(* IEC 61131-3 sources: kns-pump-station/tests/POUs/Station/FB_StationCore_Test, 49 files *)

(* ---- AlarmIdCommandsResultAndClear.method.decl.st ---- *)
// 08 §14 вопрос 1: номера udiAckId, udiShelveId, udiUnshelveId — команда засчитывается, номер сбрасывается,
// результат — по ответу сводки
METHOD PRIVATE AlarmIdCommandsResultAndClear
VAR
    fbDut        : FB_StationCore;                    // ФБ под тестом
    fbTime       : PL.FB_FakeTime;                    // подменное время, старт 1 ч
    fbSink       : FB_FakeEventSink;                  // подменный журнал
    afbPump      : ARRAY[1..3] OF FB_FakeMotorVfd;    // подменные насосы: доступны, Auto, стоят
    stCmd        : ST_StationCmd;                     // GVL_Station.stStationCmd
    stCfgPersist : ST_StationCfg;                     // GVL_Persist.stStationCfg
    stCfgLkg     : ST_StationCfg;                     // GVL_Station.stCfgLkg
    stRetain     : ST_StationRetain;                  // GVL_Persist.stStationRetain
    fbPid        : PL.FB_PID;                         // GVL_Station.fbLIC101
    stPidCmd     : PL.ST_PidCmd;                      // GVL_Station.stLIC101Cmd
    stPidCfg     : PL.ST_PidCfg;                      // GVL_Persist.stLIC101Cfg
    stPidRetain  : PL.ST_DeviceRetain;                // GVL_Persist.stLIC101Retain
    fbAlarms     : FB_StationAlarms;                  // GVL_Station.fbAlarms
END_VAR

(* ---- ApplyProjectCfgChecksProjectLevelLimits.method.decl.st ---- *)
// 04 §18.3, DESIGN 6.15: «Применить уставки проекта» при LT101 L, перенастроенной наладчиком (1,1 м, станция —
// останов 1,2 м). PRG_Devices восстанавливает L/H LT101 уставок проекта в том же цикле, но после станции: уставки
// по умолчанию (останов 1,00 м) проверяются по L/H проекта (0,8 / 3,5 м). В цикле команды нет ложной ошибки уставок
// (NE 107 «функциональная проверка»), действующей становится копия по умолчанию, событие 101017 — одно, со значением 0
METHOD PRIVATE ApplyProjectCfgChecksProjectLevelLimits
VAR
    fbDut        : FB_StationCore;                    // ФБ под тестом
    fbTime       : PL.FB_FakeTime;                    // подменное время, старт 1 ч
    fbSink       : FB_FakeEventSink;                  // подменный журнал
    afbPump      : ARRAY[1..3] OF FB_FakeMotorVfd;    // подменные насосы: доступны, Auto, стоят
    stCmd        : ST_StationCmd;                     // GVL_Station.stStationCmd
    stCfgPersist : ST_StationCfg;                     // GVL_Persist.stStationCfg
    stCfgLkg     : ST_StationCfg;                     // GVL_Station.stCfgLkg
    stRetain     : ST_StationRetain;                  // GVL_Persist.stStationRetain
    fbPid        : PL.FB_PID;                         // GVL_Station.fbLIC101
    stPidCmd     : PL.ST_PidCmd;                      // GVL_Station.stLIC101Cmd
    stPidCfg     : PL.ST_PidCfg;                      // GVL_Persist.stLIC101Cfg
    stPidRetain  : PL.ST_DeviceRetain;                // GVL_Persist.stLIC101Retain
    fbAlarms     : FB_StationAlarms;                  // GVL_Station.fbAlarms
END_VAR

(* ---- ApplyProjectCfgRestoresDefaults.method.decl.st ---- *)
// 04 §18.3: «Применить уставки проекта» возвращает уставки станции и LIC101 к значениям GVL_StationDefaults
METHOD PRIVATE ApplyProjectCfgRestoresDefaults
VAR
    fbDut        : FB_StationCore;                    // ФБ под тестом
    fbTime       : PL.FB_FakeTime;                    // подменное время, старт 1 ч
    fbSink       : FB_FakeEventSink;                  // подменный журнал
    afbPump      : ARRAY[1..3] OF FB_FakeMotorVfd;    // подменные насосы: доступны, Auto, стоят
    stCmd        : ST_StationCmd;                     // GVL_Station.stStationCmd
    stCfgPersist : ST_StationCfg;                     // GVL_Persist.stStationCfg
    stCfgLkg     : ST_StationCfg;                     // GVL_Station.stCfgLkg
    stRetain     : ST_StationRetain;                  // GVL_Persist.stStationRetain
    fbPid        : PL.FB_PID;                         // GVL_Station.fbLIC101
    stPidCmd     : PL.ST_PidCmd;                      // GVL_Station.stLIC101Cmd
    stPidCfg     : PL.ST_PidCfg;                      // GVL_Persist.stLIC101Cfg
    stPidRetain  : PL.ST_DeviceRetain;                // GVL_Persist.stLIC101Retain
    fbAlarms     : FB_StationAlarms;                  // GVL_Station.fbAlarms
END_VAR

(* ---- AtsReplacesFaultedLead.method.decl.st ---- *)
// 04 §9, PMI-12, PMI-13: отказ ведущего — замена в том же цикле, событие 101006, KNS1.ATS
METHOD PRIVATE AtsReplacesFaultedLead
VAR
    fbDut        : FB_StationCore;                    // ФБ под тестом
    fbTime       : PL.FB_FakeTime;                    // подменное время, старт 1 ч
    fbSink       : FB_FakeEventSink;                  // подменный журнал
    afbPump      : ARRAY[1..3] OF FB_FakeMotorVfd;    // подменные насосы: доступны, Auto, стоят
    stCmd        : ST_StationCmd;                     // GVL_Station.stStationCmd
    stCfgPersist : ST_StationCfg;                     // GVL_Persist.stStationCfg
    stCfgLkg     : ST_StationCfg;                     // GVL_Station.stCfgLkg
    stRetain     : ST_StationRetain;                  // GVL_Persist.stStationRetain
    fbPid        : PL.FB_PID;                         // GVL_Station.fbLIC101
    stPidCmd     : PL.ST_PidCmd;                      // GVL_Station.stLIC101Cmd
    stPidCfg     : PL.ST_PidCfg;                      // GVL_Persist.stLIC101Cfg
    stPidRetain  : PL.ST_DeviceRetain;                // GVL_Persist.stLIC101Retain
    fbAlarms     : FB_StationAlarms;                  // GVL_Station.fbAlarms
END_VAR

(* ---- CommandPulsesClearedAndCounted.method.decl.st ---- *)
// 04 §19.2, контракт 2.1: импульсы и номера команд сбрасываются в том же цикле, uiCmdSeq растёт на число команд,
// eCmdResult — последней; события 101001, 101022, 101023
METHOD PRIVATE CommandPulsesClearedAndCounted
VAR
    fbDut        : FB_StationCore;                    // ФБ под тестом
    fbTime       : PL.FB_FakeTime;                    // подменное время, старт 1 ч
    fbSink       : FB_FakeEventSink;                  // подменный журнал
    afbPump      : ARRAY[1..3] OF FB_FakeMotorVfd;    // подменные насосы: доступны, Auto, стоят
    stCmd        : ST_StationCmd;                     // GVL_Station.stStationCmd
    stCfgPersist : ST_StationCfg;                     // GVL_Persist.stStationCfg
    stCfgLkg     : ST_StationCfg;                     // GVL_Station.stCfgLkg
    stRetain     : ST_StationRetain;                  // GVL_Persist.stStationRetain
    fbPid        : PL.FB_PID;                         // GVL_Station.fbLIC101
    stPidCmd     : PL.ST_PidCmd;                      // GVL_Station.stLIC101Cmd
    stPidCfg     : PL.ST_PidCfg;                      // GVL_Persist.stLIC101Cfg
    stPidRetain  : PL.ST_DeviceRetain;                // GVL_Persist.stLIC101Retain
    fbAlarms     : FB_StationAlarms;                  // GVL_Station.fbAlarms
    uiSeq0       : UINT;                              // счётчик команд до
END_VAR

(* ---- Cycle.method.decl.st ---- *)
// Помощник: uiSteps шагов времени tStep с вызовом ядра станции и всеми данными GVL_Station и
// GVL_Persist. xPlant — подменные насосы в Auto следуют запросам и общему заданию частоты
// (видно со следующего шага): работают, если запрошены, доступны и без отказа
METHOD PRIVATE Cycle
VAR_IN_OUT
    fbDut        : FB_StationCore;                    // ФБ под тестом
    fbTime       : PL.FB_FakeTime;                    // подменное время
    stCmd        : ST_StationCmd;                     // команды
    stCfgPersist : ST_StationCfg;                     // записанные уставки
    stCfgLkg     : ST_StationCfg;                     // действующая копия
    stRetain     : ST_StationRetain;                  // режим, способ
    fbPid        : PL.FB_PID;                         // LIC101
    stPidCmd     : PL.ST_PidCmd;                      // команды LIC101
    stPidCfg     : PL.ST_PidCfg;                      // уставки LIC101
    stPidRetain  : PL.ST_DeviceRetain;                // режим LIC101
    fbAlarms     : FB_StationAlarms;                  // тревоги станции
    afbPump      : ARRAY[1..3] OF FB_FakeMotorVfd;    // подменные насосы
END_VAR
VAR_INPUT
    tStep   : TIME;                                   // шаг времени
    uiSteps : UINT;                                   // шагов
    xPlant  : BOOL;                                   // насосы следуют запросам
END_VAR
VAR
    uiStep : UINT;                                    // номер шага
    uiIdx  : UINT;                                    // насос
END_VAR

(* ---- Cycle.method.impl.st ---- *)
FOR uiStep := 1 TO uiSteps DO
    fbTime.Advance(tStep := tStep);
    // сохранённая копия LKG — та же переменная, что и действующая: перезапуск ПЛК эти тесты не моделируют
    fbDut(itfTime := fbTime, stCmd := stCmd, stCfgPersist := stCfgPersist, stCfgLkg := stCfgLkg,
          stCfgLkgRetain := stCfgLkg, stRetain := stRetain, fbLIC101 := fbPid, stLIC101Cmd := stPidCmd,
          stLIC101Cfg := stPidCfg, stLIC101Retain := stPidRetain, fbAlarms := fbAlarms);
    IF xPlant THEN
        FOR uiIdx := 1 TO 3 DO
            IF afbPump[uiIdx].eMode = PL.E_DeviceMode.Auto THEN
                afbPump[uiIdx].xRunning := fbDut.axRun[uiIdx] AND afbPump[uiIdx].xAvailable
                                           AND NOT afbPump[uiIdx].xFault;
                afbPump[uiIdx].xSpeedAuto := afbPump[uiIdx].xRunning;
                afbPump[uiIdx].rSpeedRef := SEL(afbPump[uiIdx].xRunning, 0.0, fbDut.rSpeedSp_pct);
                afbPump[uiIdx].rSpeedAct := afbPump[uiIdx].rSpeedRef;
            END_IF
        END_FOR
    END_IF
END_FOR

(* ---- DryRunReleaseNoNoresStepFlicker.method.decl.st ---- *)
// 04 §7.4, §10.1, §15, PMI-22: выбран ПИД, сухой ход по LL дольше выдержек KNS1.NORES и KNS1.STEP (10 с) —
// обе подавлены (насосы заблокированы защитой станции). Насос видит снятие блокировки в своём вызове — после
// станции: в цикле снятия сухого хода насосы ещё недоступны, ПИД не готов. Ни NORES (High: сирена, K1), ни STEP
// не мелькают: выдержка появления отсчитывается заново после снятия подавления; затем снова ПИД
METHOD PRIVATE DryRunReleaseNoNoresStepFlicker
VAR
    fbDut        : FB_StationCore;                    // ФБ под тестом
    fbTime       : PL.FB_FakeTime;                    // подменное время, старт 1 ч
    fbSink       : FB_FakeEventSink;                  // подменный журнал
    afbPump      : ARRAY[1..3] OF FB_FakeMotorVfd;    // подменные насосы: доступны, Auto, стоят
    stCmd        : ST_StationCmd;                     // GVL_Station.stStationCmd
    stCfgPersist : ST_StationCfg;                     // GVL_Persist.stStationCfg
    stCfgLkg     : ST_StationCfg;                     // GVL_Station.stCfgLkg
    stRetain     : ST_StationRetain;                  // GVL_Persist.stStationRetain
    fbPid        : PL.FB_PID;                         // GVL_Station.fbLIC101
    stPidCmd     : PL.ST_PidCmd;                      // GVL_Station.stLIC101Cmd
    stPidCfg     : PL.ST_PidCfg;                      // GVL_Persist.stLIC101Cfg
    stPidRetain  : PL.ST_DeviceRetain;                // GVL_Persist.stLIC101Retain
    fbAlarms     : FB_StationAlarms;                  // GVL_Station.fbAlarms
    itfNores     : PL.I_Alarm;                        // KNS1.NORES через интерфейс
    itfStep      : PL.I_Alarm;                        // KNS1.STEP через интерфейс
    uiIdx        : UINT;                              // насос
    uiStep       : UINT;                              // шаг
    xFlicker     : BOOL;                              // NORES или STEP были неквитированными хотя бы в одном цикле
END_VAR

(* ---- DryRunReleaseNoNoresStepFlicker.method.impl.st ---- *)
coUnit.TEST('StationCore_DryRunReleaseNoNoresStepFlicker_A7_A10_A15_PMI22');

stPidCfg := GVL_StationDefaults.stLIC101Cfg;
stRetain.eMode := E_StationMode.Auto;
stRetain.eMethod := E_ControlMethod.LevelPid;
stPidRetain.eRemoteMode := PL.E_DeviceMode.Auto;
fbDut.aitfPump[1] := afbPump[1];
fbDut.aitfPump[2] := afbPump[2];
fbDut.aitfPump[3] := afbPump[3];
fbDut.axCommOk[1] := TRUE;
fbDut.axCommOk[2] := TRUE;
fbDut.axCommOk[3] := TRUE;
fbDut.itfEvents := fbSink;
fbDut.rLevel_m := 1.2;
fbDut.xLevelValid := TRUE;
fbDut.eLevelNe107 := PL.E_Ne107Status.Good;
fbDut.rLvlL_m := 0.8;
fbDut.rLvlH_m := 3.5;
fbDut.xPowerOk := TRUE;
Cycle(fbDut := fbDut, fbTime := fbTime, stCmd := stCmd, stCfgPersist := stCfgPersist, stCfgLkg := stCfgLkg,
      stRetain := stRetain, fbPid := fbPid, stPidCmd := stPidCmd, stPidCfg := stPidCfg,
      stPidRetain := stPidRetain, fbAlarms := fbAlarms, afbPump := afbPump, tStep := T#100MS, uiSteps := 110,
      xPlant := TRUE);

AssertTrue(Condition := fbDut.stSts.eControlAct = E_ControlAct.LevelPid, Message := 'LevelPid before dry run');
// LL по уровнемеру: сухой ход 20 с; насос недоступен с цикла после блокировки (как устройство после станции)
fbDut.rLevel_m := 0.45;
fbDut.xLevelL := TRUE;
fbDut.xLevelLL := TRUE;
FOR uiStep := 1 TO 200 DO
    Cycle(fbDut := fbDut, fbTime := fbTime, stCmd := stCmd, stCfgPersist := stCfgPersist, stCfgLkg := stCfgLkg,
          stRetain := stRetain, fbPid := fbPid, stPidCmd := stPidCmd, stPidCfg := stPidCfg,
          stPidRetain := stPidRetain, fbAlarms := fbAlarms, afbPump := afbPump, tStep := T#100MS, uiSteps := 1,
          xPlant := TRUE);
    FOR uiIdx := 1 TO 3 DO
        afbPump[uiIdx].xAvailable := fbDut.awInterlock[uiIdx] = 0;
    END_FOR
END_FOR

AssertTrue(Condition := fbDut.stSts.eControlAct = E_ControlAct.DryRunStop, Message := 'DryRunStop');
itfNores := fbAlarms.GetAlarm(uiIndex := E_StationAlarm.NORES - 1);
itfStep := fbAlarms.GetAlarm(uiIndex := E_StationAlarm.STEP - 1);
AssertTrue(Condition := itfNores.State = PL.E_AlarmState.SuppressedByDesign, Message := 'dry run: NORES suppressed');
AssertTrue(Condition := itfStep.State = PL.E_AlarmState.SuppressedByDesign, Message := 'dry run: STEP suppressed');
// уровень выше L: сухой ход снят
fbDut.rLevel_m := 1.0;
fbDut.xLevelL := FALSE;
fbDut.xLevelLL := FALSE;
xFlicker := FALSE;
FOR uiStep := 1 TO 150 DO
    Cycle(fbDut := fbDut, fbTime := fbTime, stCmd := stCmd, stCfgPersist := stCfgPersist, stCfgLkg := stCfgLkg,
          stRetain := stRetain, fbPid := fbPid, stPidCmd := stPidCmd, stPidCfg := stPidCfg,
          stPidRetain := stPidRetain, fbAlarms := fbAlarms, afbPump := afbPump, tStep := T#100MS, uiSteps := 1,
          xPlant := TRUE);
    IF uiStep = 1 THEN
        AssertEquals_UINT(Expected := 0, Actual := fbDut.stSts.uiPumpsAvailable,
                          Message := 'release cycle: pumps still interlocked');
    END_IF
    xFlicker := xFlicker OR (fbDut.stSts.wAlmUnack AND 16#0088) <> 0;
    FOR uiIdx := 1 TO 3 DO
        afbPump[uiIdx].xAvailable := fbDut.awInterlock[uiIdx] = 0;
    END_FOR
END_FOR

AssertFalse(Condition := xFlicker, Message := 'no unacked KNS1.NORES or KNS1.STEP on dry run release');
AssertTrue(Condition := itfNores.State = PL.E_AlarmState.Normal, Message := 'NORES normal');
AssertTrue(Condition := itfStep.State = PL.E_AlarmState.Normal, Message := 'STEP normal');
AssertTrue(Condition := fbDut.stSts.eControlAct = E_ControlAct.LevelPid, Message := 'LevelPid after dry run');

coUnit.TEST_FINISHED();

(* ---- DryRunStopSuppressesNoReserve.method.decl.st ---- *)
// 04 §10.1, §11, §15, PMI-21: откачка по поплавкам до LS103 — сухой ход блокирует все насосы (Available = FALSE).
// Насосы стоят по защите станции, а не из-за отказов: KNS1.NORES подавлена (дубль KNS1.DRY, иначе High-тревога и
// обесточенное K1 в каждом цикле откачки по поплавкам)
METHOD PRIVATE DryRunStopSuppressesNoReserve
VAR
    fbDut        : FB_StationCore;                    // ФБ под тестом
    fbTime       : PL.FB_FakeTime;                    // подменное время, старт 1 ч
    fbSink       : FB_FakeEventSink;                  // подменный журнал
    afbPump      : ARRAY[1..3] OF FB_FakeMotorVfd;    // подменные насосы: доступны, Auto, стоят
    stCmd        : ST_StationCmd;                     // GVL_Station.stStationCmd
    stCfgPersist : ST_StationCfg;                     // GVL_Persist.stStationCfg
    stCfgLkg     : ST_StationCfg;                     // GVL_Station.stCfgLkg
    stRetain     : ST_StationRetain;                  // GVL_Persist.stStationRetain
    fbPid        : PL.FB_PID;                         // GVL_Station.fbLIC101
    stPidCmd     : PL.ST_PidCmd;                      // GVL_Station.stLIC101Cmd
    stPidCfg     : PL.ST_PidCfg;                      // GVL_Persist.stLIC101Cfg
    stPidRetain  : PL.ST_DeviceRetain;                // GVL_Persist.stLIC101Retain
    fbAlarms     : FB_StationAlarms;                  // GVL_Station.fbAlarms
    itfAlm       : PL.I_Alarm;                        // тревога через интерфейс
    uiIdx        : UINT;                              // насос
END_VAR

(* ---- DryRunStopSuppressesNoReserve.method.impl.st ---- *)
coUnit.TEST('StationCore_DryRunStopSuppressesNoReserve_A10_A11_A15_PMI21');

stPidCfg := GVL_StationDefaults.stLIC101Cfg;
stRetain.eMode := E_StationMode.Auto;
fbDut.aitfPump[1] := afbPump[1];
fbDut.aitfPump[2] := afbPump[2];
fbDut.aitfPump[3] := afbPump[3];
fbDut.axCommOk[1] := TRUE;
fbDut.axCommOk[2] := TRUE;
fbDut.axCommOk[3] := TRUE;
fbDut.itfEvents := fbSink;
fbDut.rLevel_m := 1.2;
fbDut.xLevelValid := TRUE;
fbDut.eLevelNe107 := PL.E_Ne107Status.Good;
fbDut.rLvlL_m := 0.8;
fbDut.rLvlH_m := 3.5;
fbDut.xPowerOk := TRUE;
Cycle(fbDut := fbDut, fbTime := fbTime, stCmd := stCmd, stCfgPersist := stCfgPersist, stCfgLkg := stCfgLkg,
      stRetain := stRetain, fbPid := fbPid, stPidCmd := stPidCmd, stPidCfg := stPidCfg,
      stPidRetain := stPidRetain, fbAlarms := fbAlarms, afbPump := afbPump, tStep := T#100MS, uiSteps := 110,
      xPlant := TRUE);

// отказ LT101, LS102: откачка всеми насосами
fbDut.xLevelValid := FALSE;
fbDut.xFloatHigh := TRUE;
Cycle(fbDut := fbDut, fbTime := fbTime, stCmd := stCmd, stCfgPersist := stCfgPersist, stCfgLkg := stCfgLkg,
      stRetain := stRetain, fbPid := fbPid, stPidCmd := stPidCmd, stPidCfg := stPidCfg,
      stPidRetain := stPidRetain, fbAlarms := fbAlarms, afbPump := afbPump, tStep := T#100MS, uiSteps := 110,
      xPlant := TRUE);

AssertTrue(Condition := afbPump[1].xRunning AND afbPump[2].xRunning AND afbPump[3].xRunning, Message := 'pumping');
// уровень у LS103: сухой ход, блокировка всех насосов — устройства недоступны и стоят
fbDut.xFloatHigh := FALSE;
fbDut.xFloatDry := TRUE;
Cycle(fbDut := fbDut, fbTime := fbTime, stCmd := stCmd, stCfgPersist := stCfgPersist, stCfgLkg := stCfgLkg,
      stRetain := stRetain, fbPid := fbPid, stPidCmd := stPidCmd, stPidCfg := stPidCfg,
      stPidRetain := stPidRetain, fbAlarms := fbAlarms, afbPump := afbPump, tStep := T#100MS, uiSteps := 1,
      xPlant := TRUE);

AssertTrue(Condition := (fbDut.awInterlock[1] AND GVL_Const.KNS_ILK_DRY_RUN) <> 0, Message := 'dry run interlock');
FOR uiIdx := 1 TO 3 DO
    afbPump[uiIdx].xAvailable := FALSE;
END_FOR
Cycle(fbDut := fbDut, fbTime := fbTime, stCmd := stCmd, stCfgPersist := stCfgPersist, stCfgLkg := stCfgLkg,
      stRetain := stRetain, fbPid := fbPid, stPidCmd := stPidCmd, stPidCfg := stPidCfg,
      stPidRetain := stPidRetain, fbAlarms := fbAlarms, afbPump := afbPump, tStep := T#100MS, uiSteps := 200,
      xPlant := TRUE);

AssertTrue(Condition := fbDut.stSts.eControlAct = E_ControlAct.DryRunStop, Message := 'DryRunStop');
AssertEquals_UINT(Expected := 0, Actual := fbDut.stSts.uiPumpsAvailable, Message := 'no pump available');
itfAlm := fbAlarms.GetAlarm(uiIndex := E_StationAlarm.NORES - 1);
AssertTrue(Condition := itfAlm.State = PL.E_AlarmState.SuppressedByDesign, Message := 'NORES suppressed by dry run');
AssertEquals_WORD(Expected := 0, Actual := fbDut.stSts.wAlmActive AND 16#0004, Message := 'no LACK');
AssertEquals_WORD(Expected := 0, Actual := fbDut.stSts.wAlmUnack AND 16#000C, Message := 'no LACK, NORES unacked');
AssertEquals_WORD(Expected := 0, Actual := fbDut.stSts.wState AND GVL_Const.STN_ST_NO_RESERVE,
                  Message := 'wState: no reserve bit clear');

coUnit.TEST_FINISHED();

(* ---- EmergencyRequiresAllAtFullSpeed.method.decl.st ---- *)
// 04 §10.2, PMI-20: аварийный уровень в «Автомате» — требуются все три насоса, задание 100 %, KNS1.EHL, K1 по
// сводке
METHOD PRIVATE EmergencyRequiresAllAtFullSpeed
VAR
    fbDut        : FB_StationCore;                    // ФБ под тестом
    fbTime       : PL.FB_FakeTime;                    // подменное время, старт 1 ч
    fbSink       : FB_FakeEventSink;                  // подменный журнал
    afbPump      : ARRAY[1..3] OF FB_FakeMotorVfd;    // подменные насосы: доступны, Auto, стоят
    stCmd        : ST_StationCmd;                     // GVL_Station.stStationCmd
    stCfgPersist : ST_StationCfg;                     // GVL_Persist.stStationCfg
    stCfgLkg     : ST_StationCfg;                     // GVL_Station.stCfgLkg
    stRetain     : ST_StationRetain;                  // GVL_Persist.stStationRetain
    fbPid        : PL.FB_PID;                         // GVL_Station.fbLIC101
    stPidCmd     : PL.ST_PidCmd;                      // GVL_Station.stLIC101Cmd
    stPidCfg     : PL.ST_PidCfg;                      // GVL_Persist.stLIC101Cfg
    stPidRetain  : PL.ST_DeviceRetain;                // GVL_Persist.stLIC101Retain
    fbAlarms     : FB_StationAlarms;                  // GVL_Station.fbAlarms
END_VAR

(* ---- ExportCommandAndEvents.method.decl.st ---- *)
// 04 §16, PMI-37: xExportLog — запрос снимка; во время выгрузки отклоняется; переход в Done — событие 101019 с
// числом строк, в Error — 101020
METHOD PRIVATE ExportCommandAndEvents
VAR
    fbDut        : FB_StationCore;                    // ФБ под тестом
    fbTime       : PL.FB_FakeTime;                    // подменное время, старт 1 ч
    fbSink       : FB_FakeEventSink;                  // подменный журнал
    afbPump      : ARRAY[1..3] OF FB_FakeMotorVfd;    // подменные насосы: доступны, Auto, стоят
    stCmd        : ST_StationCmd;                     // GVL_Station.stStationCmd
    stCfgPersist : ST_StationCfg;                     // GVL_Persist.stStationCfg
    stCfgLkg     : ST_StationCfg;                     // GVL_Station.stCfgLkg
    stRetain     : ST_StationRetain;                  // GVL_Persist.stStationRetain
    fbPid        : PL.FB_PID;                         // GVL_Station.fbLIC101
    stPidCmd     : PL.ST_PidCmd;                      // GVL_Station.stLIC101Cmd
    stPidCfg     : PL.ST_PidCfg;                      // GVL_Persist.stLIC101Cfg
    stPidRetain  : PL.ST_DeviceRetain;                // GVL_Persist.stLIC101Retain
    fbAlarms     : FB_StationAlarms;                  // GVL_Station.fbAlarms
END_VAR

(* ---- FloatModeStartsAllOnLs102.method.decl.st ---- *)
// 04 §11, PMI-21, PMI-25: LT101 недостоверен — Float; LS102 — все насосы, 100 %; KNS1.EHL и KNS1.DRY подавлены,
// KNS1.FLOAT активна
METHOD PRIVATE FloatModeStartsAllOnLs102
VAR
    fbDut        : FB_StationCore;                    // ФБ под тестом
    fbTime       : PL.FB_FakeTime;                    // подменное время, старт 1 ч
    fbSink       : FB_FakeEventSink;                  // подменный журнал
    afbPump      : ARRAY[1..3] OF FB_FakeMotorVfd;    // подменные насосы: доступны, Auto, стоят
    stCmd        : ST_StationCmd;                     // GVL_Station.stStationCmd
    stCfgPersist : ST_StationCfg;                     // GVL_Persist.stStationCfg
    stCfgLkg     : ST_StationCfg;                     // GVL_Station.stCfgLkg
    stRetain     : ST_StationRetain;                  // GVL_Persist.stStationRetain
    fbPid        : PL.FB_PID;                         // GVL_Station.fbLIC101
    stPidCmd     : PL.ST_PidCmd;                      // GVL_Station.stLIC101Cmd
    stPidCfg     : PL.ST_PidCfg;                      // GVL_Persist.stLIC101Cfg
    stPidRetain  : PL.ST_DeviceRetain;                // GVL_Persist.stLIC101Retain
    fbAlarms     : FB_StationAlarms;                  // GVL_Station.fbAlarms
    itfAlm       : PL.I_Alarm;                        // тревога через интерфейс
END_VAR

(* ---- FlowAlarmsSuppressedUntilSettled.method.decl.st ---- *)
// DESIGN 7, шаг 12: тревоги L/LL PT201 и L FT202 подавлены, пока ни один насос не работает дольше STN_FLOW_SETTLE
// = 20 с
METHOD PRIVATE FlowAlarmsSuppressedUntilSettled
VAR
    fbDut        : FB_StationCore;                    // ФБ под тестом
    fbTime       : PL.FB_FakeTime;                    // подменное время, старт 1 ч
    fbSink       : FB_FakeEventSink;                  // подменный журнал
    afbPump      : ARRAY[1..3] OF FB_FakeMotorVfd;    // подменные насосы: доступны, Auto, стоят
    stCmd        : ST_StationCmd;                     // GVL_Station.stStationCmd
    stCfgPersist : ST_StationCfg;                     // GVL_Persist.stStationCfg
    stCfgLkg     : ST_StationCfg;                     // GVL_Station.stCfgLkg
    stRetain     : ST_StationRetain;                  // GVL_Persist.stStationRetain
    fbPid        : PL.FB_PID;                         // GVL_Station.fbLIC101
    stPidCmd     : PL.ST_PidCmd;                      // GVL_Station.stLIC101Cmd
    stPidCfg     : PL.ST_PidCfg;                      // GVL_Persist.stLIC101Cfg
    stPidRetain  : PL.ST_DeviceRetain;                // GVL_Persist.stLIC101Retain
    fbAlarms     : FB_StationAlarms;                  // GVL_Station.fbAlarms
END_VAR

(* ---- LackSuppressesNoReserve.method.decl.st ---- *)
// 04 §15, PMI-17: недостаточно насосов — KNS1.LACK через 10 с, KNS1.NORES подавлена; NE 107 станции — Failure
METHOD PRIVATE LackSuppressesNoReserve
VAR
    fbDut        : FB_StationCore;                    // ФБ под тестом
    fbTime       : PL.FB_FakeTime;                    // подменное время, старт 1 ч
    fbSink       : FB_FakeEventSink;                  // подменный журнал
    afbPump      : ARRAY[1..3] OF FB_FakeMotorVfd;    // подменные насосы: доступны, Auto, стоят
    stCmd        : ST_StationCmd;                     // GVL_Station.stStationCmd
    stCfgPersist : ST_StationCfg;                     // GVL_Persist.stStationCfg
    stCfgLkg     : ST_StationCfg;                     // GVL_Station.stCfgLkg
    stRetain     : ST_StationRetain;                  // GVL_Persist.stStationRetain
    fbPid        : PL.FB_PID;                         // GVL_Station.fbLIC101
    stPidCmd     : PL.ST_PidCmd;                      // GVL_Station.stLIC101Cmd
    stPidCfg     : PL.ST_PidCfg;                      // GVL_Persist.stLIC101Cfg
    stPidRetain  : PL.ST_DeviceRetain;                // GVL_Persist.stLIC101Retain
    fbAlarms     : FB_StationAlarms;                  // GVL_Station.fbAlarms
    itfAlm       : PL.I_Alarm;                        // тревога через интерфейс
END_VAR

(* ---- LkgRejectsInvalidCfg.method.decl.st ---- *)
// 04 §18.3, PMI-08: корректная уставка принимается (событие 101017 с номером параметра 8), неверная не применяется
// — бит wCfgErr, работа по последней корректной копии
METHOD PRIVATE LkgRejectsInvalidCfg
VAR
    fbDut        : FB_StationCore;                    // ФБ под тестом
    fbTime       : PL.FB_FakeTime;                    // подменное время, старт 1 ч
    fbSink       : FB_FakeEventSink;                  // подменный журнал
    afbPump      : ARRAY[1..3] OF FB_FakeMotorVfd;    // подменные насосы: доступны, Auto, стоят
    stCmd        : ST_StationCmd;                     // GVL_Station.stStationCmd
    stCfgPersist : ST_StationCfg;                     // GVL_Persist.stStationCfg
    stCfgLkg     : ST_StationCfg;                     // GVL_Station.stCfgLkg
    stRetain     : ST_StationRetain;                  // GVL_Persist.stStationRetain
    fbPid        : PL.FB_PID;                         // GVL_Station.fbLIC101
    stPidCmd     : PL.ST_PidCmd;                      // GVL_Station.stLIC101Cmd
    stPidCfg     : PL.ST_PidCfg;                      // GVL_Persist.stLIC101Cfg
    stPidRetain  : PL.ST_DeviceRetain;                // GVL_Persist.stLIC101Retain
    fbAlarms     : FB_StationAlarms;                  // GVL_Station.fbAlarms
END_VAR

(* ---- LkgRestoredAfterRestart.method.decl.st ---- *)
// 04 §18.3, PMI-08, PMI-35: последняя корректная копия уставок переживает перезапуск ПЛК. Корректная правка
// (задание 1,8 м) принята и сохранена в энергонезависимой копии LKG, неверная (2,5 м) осталась в записанных
// уставках; после перезапуска (новый экземпляр ядра, GVL_Station.stCfgLkg — умолчания) станция работает по
// сохранённой копии 1,8 м, а не по уставкам проекта; событие 101017 при старте не пишется
METHOD PRIVATE LkgRestoredAfterRestart
VAR
    fbTime         : PL.FB_FakeTime;                  // подменное время, старт 1 ч
    afbPump        : ARRAY[1..3] OF FB_FakeMotorVfd;  // подменные насосы: доступны, Auto, стоят
    // энергонезависимые данные (GVL_Persist): переживают перезапуск
    stCfgPersist   : ST_StationCfg;                   // GVL_Persist.stStationCfg
    stCfgLkgRetain : ST_StationCfg;                   // GVL_Persist.stStationCfgLkg
    stRetain       : ST_StationRetain;                // GVL_Persist.stStationRetain
    stPidCfg       : PL.ST_PidCfg;                    // GVL_Persist.stLIC101Cfg
    stPidRetain    : PL.ST_DeviceRetain;              // GVL_Persist.stLIC101Retain
END_VAR
VAR_INST
    // до перезапуска
    fbDutBefore    : FB_StationCore;                  // ядро до перезапуска
    fbSinkBefore   : FB_FakeEventSink;                // журнал до перезапуска
    stCmdBefore    : ST_StationCmd;                   // GVL_Station.stStationCmd
    stLkgBefore    : ST_StationCfg;                   // GVL_Station.stCfgLkg
    fbPidBefore    : PL.FB_PID;                       // GVL_Station.fbLIC101
    stPidCmdBefore : PL.ST_PidCmd;                    // GVL_Station.stLIC101Cmd
    fbAlmBefore    : FB_StationAlarms;                // GVL_Station.fbAlarms
    // после перезапуска: обычные переменные снова с умолчаниями
    fbDutAfter     : FB_StationCore;                  // ядро после перезапуска
    fbSinkAfter    : FB_FakeEventSink;                // журнал после перезапуска
    stCmdAfter     : ST_StationCmd;
    stLkgAfter     : ST_StationCfg;
    fbPidAfter     : PL.FB_PID;
    stPidCmdAfter  : PL.ST_PidCmd;
    fbAlmAfter     : FB_StationAlarms;
END_VAR

(* ---- ManualDryRunInterlocksAllPumps.method.decl.st ---- *)
// 04 §10.1, PMI-18: в «Ручном» запросов нет, но сухой ход по LL блокирует все насосы (KNS_ILK_DRY_RUN), тревога
// KNS1.DRY
METHOD PRIVATE ManualDryRunInterlocksAllPumps
VAR
    fbDut        : FB_StationCore;                    // ФБ под тестом
    fbTime       : PL.FB_FakeTime;                    // подменное время, старт 1 ч
    fbSink       : FB_FakeEventSink;                  // подменный журнал
    afbPump      : ARRAY[1..3] OF FB_FakeMotorVfd;    // подменные насосы: доступны, Auto, стоят
    stCmd        : ST_StationCmd;                     // GVL_Station.stStationCmd
    stCfgPersist : ST_StationCfg;                     // GVL_Persist.stStationCfg
    stCfgLkg     : ST_StationCfg;                     // GVL_Station.stCfgLkg
    stRetain     : ST_StationRetain;                  // GVL_Persist.stStationRetain
    fbPid        : PL.FB_PID;                         // GVL_Station.fbLIC101
    stPidCmd     : PL.ST_PidCmd;                      // GVL_Station.stLIC101Cmd
    stPidCfg     : PL.ST_PidCfg;                      // GVL_Persist.stLIC101Cfg
    stPidRetain  : PL.ST_DeviceRetain;                // GVL_Persist.stLIC101Retain
    fbAlarms     : FB_StationAlarms;                  // GVL_Station.fbAlarms
END_VAR

(* ---- ManualFloatModeKeepsEhlDry.method.decl.st ---- *)
// 04 §3.1, §10.2, §11, §15: станция в «Ручном», LT101 отказал. Управления по поплавкам в «Ручном» нет (насосы
// автоматика не пускает), поэтому KNS1.EHL (Critical) по LS102 и KNS1.DRY по LS103 не подавляются: подавление
// «режим по поплавкам» действует только в «Автомате», где срабатывания поплавков — штатные точки управления
METHOD PRIVATE ManualFloatModeKeepsEhlDry
VAR
    fbDut        : FB_StationCore;                    // ФБ под тестом
    fbTime       : PL.FB_FakeTime;                    // подменное время, старт 1 ч
    fbSink       : FB_FakeEventSink;                  // подменный журнал
    afbPump      : ARRAY[1..3] OF FB_FakeMotorVfd;    // подменные насосы: доступны, Auto, стоят
    stCmd        : ST_StationCmd;                     // GVL_Station.stStationCmd
    stCfgPersist : ST_StationCfg;                     // GVL_Persist.stStationCfg
    stCfgLkg     : ST_StationCfg;                     // GVL_Station.stCfgLkg
    stRetain     : ST_StationRetain;                  // GVL_Persist.stStationRetain
    fbPid        : PL.FB_PID;                         // GVL_Station.fbLIC101
    stPidCmd     : PL.ST_PidCmd;                      // GVL_Station.stLIC101Cmd
    stPidCfg     : PL.ST_PidCfg;                      // GVL_Persist.stLIC101Cfg
    stPidRetain  : PL.ST_DeviceRetain;                // GVL_Persist.stLIC101Retain
    fbAlarms     : FB_StationAlarms;                  // GVL_Station.fbAlarms
    itfEhl       : PL.I_Alarm;                        // KNS1.EHL через интерфейс
    itfDry       : PL.I_Alarm;                        // KNS1.DRY через интерфейс
END_VAR

(* ---- ManualToAutoAdoptsRunningPump.method.decl.st ---- *)
// 04 §3.2, PMI-30: «Ручной» → «Автомат» при работающем насосе — в том же цикле запрос ему (без останова), насосам
// — RequestMode(Auto), задание частоты следило за насосом
METHOD PRIVATE ManualToAutoAdoptsRunningPump
VAR
    fbDut        : FB_StationCore;                    // ФБ под тестом
    fbTime       : PL.FB_FakeTime;                    // подменное время, старт 1 ч
    fbSink       : FB_FakeEventSink;                  // подменный журнал
    afbPump      : ARRAY[1..3] OF FB_FakeMotorVfd;    // подменные насосы: доступны, Auto, стоят
    stCmd        : ST_StationCmd;                     // GVL_Station.stStationCmd
    stCfgPersist : ST_StationCfg;                     // GVL_Persist.stStationCfg
    stCfgLkg     : ST_StationCfg;                     // GVL_Station.stCfgLkg
    stRetain     : ST_StationRetain;                  // GVL_Persist.stStationRetain
    fbPid        : PL.FB_PID;                         // GVL_Station.fbLIC101
    stPidCmd     : PL.ST_PidCmd;                      // GVL_Station.stLIC101Cmd
    stPidCfg     : PL.ST_PidCfg;                      // GVL_Persist.stLIC101Cfg
    stPidRetain  : PL.ST_DeviceRetain;                // GVL_Persist.stLIC101Retain
    fbAlarms     : FB_StationAlarms;                  // GVL_Station.fbAlarms
END_VAR

(* ---- ManualToAutoStoppedPumpsNoNoresFlicker.method.decl.st ---- *)
// 04 §3.2, §15, PMI-30: «Ручной» дольше выдержки KNS1.NORES (10 с) при остановленных насосах, затем «Автомат».
// Насос выполняет запрос режима в своём вызове — после станции: в цикле входа в «Автомат» насосы ещё в Manual
// (доступных нет), подавление «Ручной» уже снято, а требуемое число 0 (KNS1.LACK нет). Тревога не мелькает
// (High: сирена, K1): выдержка появления отсчитывается заново после снятия подавления
METHOD PRIVATE ManualToAutoStoppedPumpsNoNoresFlicker
VAR
    fbDut        : FB_StationCore;                    // ФБ под тестом
    fbTime       : PL.FB_FakeTime;                    // подменное время, старт 1 ч
    fbSink       : FB_FakeEventSink;                  // подменный журнал
    afbPump      : ARRAY[1..3] OF FB_FakeMotorVfd;    // подменные насосы: доступны, Auto, стоят
    stCmd        : ST_StationCmd;                     // GVL_Station.stStationCmd
    stCfgPersist : ST_StationCfg;                     // GVL_Persist.stStationCfg
    stCfgLkg     : ST_StationCfg;                     // GVL_Station.stCfgLkg
    stRetain     : ST_StationRetain;                  // GVL_Persist.stStationRetain
    fbPid        : PL.FB_PID;                         // GVL_Station.fbLIC101
    stPidCmd     : PL.ST_PidCmd;                      // GVL_Station.stLIC101Cmd
    stPidCfg     : PL.ST_PidCfg;                      // GVL_Persist.stLIC101Cfg
    stPidRetain  : PL.ST_DeviceRetain;                // GVL_Persist.stLIC101Retain
    fbAlarms     : FB_StationAlarms;                  // GVL_Station.fbAlarms
    itfAlm       : PL.I_Alarm;                        // KNS1.NORES через интерфейс
    uiIdx        : UINT;                              // насос
    uiStep       : UINT;                              // шаг
    xFlicker     : BOOL;                              // NORES была неквитированной хотя бы в одном цикле
END_VAR

(* ---- ManualToAutoStoppedPumpsNoNoresFlicker.method.impl.st ---- *)
coUnit.TEST('StationCore_ManualToAutoStoppedPumpsNoNoresFlicker_A3_A15_PMI30');

stPidCfg := GVL_StationDefaults.stLIC101Cfg;
stRetain.eMode := E_StationMode.Auto;
fbDut.aitfPump[1] := afbPump[1];
fbDut.aitfPump[2] := afbPump[2];
fbDut.aitfPump[3] := afbPump[3];
fbDut.axCommOk[1] := TRUE;
fbDut.axCommOk[2] := TRUE;
fbDut.axCommOk[3] := TRUE;
fbDut.itfEvents := fbSink;
fbDut.rLevel_m := 1.2;
fbDut.xLevelValid := TRUE;
fbDut.eLevelNe107 := PL.E_Ne107Status.Good;
fbDut.rLvlL_m := 0.8;
fbDut.rLvlH_m := 3.5;
fbDut.xPowerOk := TRUE;
Cycle(fbDut := fbDut, fbTime := fbTime, stCmd := stCmd, stCfgPersist := stCfgPersist, stCfgLkg := stCfgLkg,
      stRetain := stRetain, fbPid := fbPid, stPidCmd := stPidCmd, stPidCfg := stPidCfg,
      stPidRetain := stPidRetain, fbAlarms := fbAlarms, afbPump := afbPump, tStep := T#100MS, uiSteps := 110,
      xPlant := TRUE);

// «Ручной»: насосы выполняют запрос в своём вызове (циклом позже станции)
stCmd.xSetManual := TRUE;
Cycle(fbDut := fbDut, fbTime := fbTime, stCmd := stCmd, stCfgPersist := stCfgPersist, stCfgLkg := stCfgLkg,
      stRetain := stRetain, fbPid := fbPid, stPidCmd := stPidCmd, stPidCfg := stPidCfg,
      stPidRetain := stPidRetain, fbAlarms := fbAlarms, afbPump := afbPump, tStep := T#100MS, uiSteps := 1,
      xPlant := TRUE);

FOR uiIdx := 1 TO 3 DO
    afbPump[uiIdx].eMode := afbPump[uiIdx].eLastModeRequest;
END_FOR
AssertTrue(Condition := afbPump[1].eMode = PL.E_DeviceMode.Manual, Message := 'pumps in Manual');
Cycle(fbDut := fbDut, fbTime := fbTime, stCmd := stCmd, stCfgPersist := stCfgPersist, stCfgLkg := stCfgLkg,
      stRetain := stRetain, fbPid := fbPid, stPidCmd := stPidCmd, stPidCfg := stPidCfg,
      stPidRetain := stPidRetain, fbAlarms := fbAlarms, afbPump := afbPump, tStep := T#100MS, uiSteps := 150,
      xPlant := TRUE);

itfAlm := fbAlarms.GetAlarm(uiIndex := E_StationAlarm.NORES - 1);
AssertTrue(Condition := itfAlm.State = PL.E_AlarmState.SuppressedByDesign, Message := 'Manual 15 s: NORES suppressed');
// «Автомат»: в этом цикле насосы ещё в Manual, со следующего — в Auto
stCmd.xSetAuto := TRUE;
xFlicker := FALSE;
FOR uiStep := 1 TO 120 DO
    Cycle(fbDut := fbDut, fbTime := fbTime, stCmd := stCmd, stCfgPersist := stCfgPersist, stCfgLkg := stCfgLkg,
          stRetain := stRetain, fbPid := fbPid, stPidCmd := stPidCmd, stPidCfg := stPidCfg,
          stPidRetain := stPidRetain, fbAlarms := fbAlarms, afbPump := afbPump, tStep := T#100MS, uiSteps := 1,
          xPlant := TRUE);
    xFlicker := xFlicker OR (fbDut.stSts.wAlmUnack AND 16#0008) <> 0;
    IF uiStep = 1 THEN
        AssertEquals_UINT(Expected := 0, Actual := fbDut.stSts.uiPumpsAvailable,
                          Message := 'Auto entry cycle: pumps still in Manual');
        FOR uiIdx := 1 TO 3 DO
            afbPump[uiIdx].eMode := afbPump[uiIdx].eLastModeRequest;
        END_FOR
    END_IF
END_FOR

AssertTrue(Condition := fbDut.stSts.eMode = E_StationMode.Auto, Message := 'station in Auto');
AssertEquals_UINT(Expected := 3, Actual := fbDut.stSts.uiPumpsAvailable, Message := 'pumps available in Auto');
AssertFalse(Condition := xFlicker, Message := 'no unacked KNS1.NORES on Auto entry');
AssertTrue(Condition := itfAlm.State = PL.E_AlarmState.Normal, Message := 'NORES normal');

coUnit.TEST_FINISHED();

(* ---- OverheatTripIsAts.method.decl.st ---- *)
// 04 §9.1, §10.4, PMI-16: перегрев обмотки ведущего — TS1n2 приходит раньше аварии ПЧ (у аварии фильтр
// tExtFaultFilter 0,2 с, у TS1n2 задержки нет). Станция блокирует насос (KNS_ILK_OVERHEAT), он останавливается и
// теряет запрос до отказа устройства — это всё равно АВР: KNS1.ATS и событие 101006 с номером замены
METHOD PRIVATE OverheatTripIsAts
VAR
    fbDut        : FB_StationCore;                    // ФБ под тестом
    fbTime       : PL.FB_FakeTime;                    // подменное время, старт 1 ч
    fbSink       : FB_FakeEventSink;                  // подменный журнал
    afbPump      : ARRAY[1..3] OF FB_FakeMotorVfd;    // подменные насосы: доступны, Auto, стоят
    stCmd        : ST_StationCmd;                     // GVL_Station.stStationCmd
    stCfgPersist : ST_StationCfg;                     // GVL_Persist.stStationCfg
    stCfgLkg     : ST_StationCfg;                     // GVL_Station.stCfgLkg
    stRetain     : ST_StationRetain;                  // GVL_Persist.stStationRetain
    fbPid        : PL.FB_PID;                         // GVL_Station.fbLIC101
    stPidCmd     : PL.ST_PidCmd;                      // GVL_Station.stLIC101Cmd
    stPidCfg     : PL.ST_PidCfg;                      // GVL_Persist.stLIC101Cfg
    stPidRetain  : PL.ST_DeviceRetain;                // GVL_Persist.stLIC101Retain
    fbAlarms     : FB_StationAlarms;                  // GVL_Station.fbAlarms
END_VAR

(* ---- PidControlsLeadSpeed.method.decl.st ---- *)
// 04 §7, PMI-04: способ ПИД, LIC101 в Auto — пуск ведущего по уровню, затем ПИД управляет: общее задание частоты =
// выход LIC101
METHOD PRIVATE PidControlsLeadSpeed
VAR
    fbDut        : FB_StationCore;                    // ФБ под тестом
    fbTime       : PL.FB_FakeTime;                    // подменное время, старт 1 ч
    fbSink       : FB_FakeEventSink;                  // подменный журнал
    afbPump      : ARRAY[1..3] OF FB_FakeMotorVfd;    // подменные насосы: доступны, Auto, стоят
    stCmd        : ST_StationCmd;                     // GVL_Station.stStationCmd
    stCfgPersist : ST_StationCfg;                     // GVL_Persist.stStationCfg
    stCfgLkg     : ST_StationCfg;                     // GVL_Station.stCfgLkg
    stRetain     : ST_StationRetain;                  // GVL_Persist.stStationRetain
    fbPid        : PL.FB_PID;                         // GVL_Station.fbLIC101
    stPidCmd     : PL.ST_PidCmd;                      // GVL_Station.stLIC101Cmd
    stPidCfg     : PL.ST_PidCfg;                      // GVL_Persist.stLIC101Cfg
    stPidRetain  : PL.ST_DeviceRetain;                // GVL_Persist.stLIC101Retain
    fbAlarms     : FB_StationAlarms;                  // GVL_Station.fbAlarms
END_VAR

(* ---- PidHandoverKeepsOutput.method.decl.st ---- *)
// 04 §7.3, §8.2 в режиме ПИД: ведущий работает непрерывно дольше tMaxContRun — передача роли резервному с
// перекрытием tOverlap; роль переходит к уже работающей замене в том же цикле, когда прежний насос теряет запрос,
// поэтому выход LIC101 и частота насосов не проваливаются ни в одном шаге передачи
METHOD PRIVATE PidHandoverKeepsOutput
VAR
    fbDut        : FB_StationCore;                    // ФБ под тестом
    fbTime       : PL.FB_FakeTime;                    // подменное время, старт 1 ч
    fbSink       : FB_FakeEventSink;                  // подменный журнал
    afbPump      : ARRAY[1..3] OF FB_FakeMotorVfd;    // подменные насосы: доступны, Auto, стоят
    stCmd        : ST_StationCmd;                     // GVL_Station.stStationCmd
    stCfgPersist : ST_StationCfg;                     // GVL_Persist.stStationCfg
    stCfgLkg     : ST_StationCfg;                     // GVL_Station.stCfgLkg
    stRetain     : ST_StationRetain;                  // GVL_Persist.stStationRetain
    fbPid        : PL.FB_PID;                         // GVL_Station.fbLIC101
    stPidCmd     : PL.ST_PidCmd;                      // GVL_Station.stLIC101Cmd
    stPidCfg     : PL.ST_PidCfg;                      // GVL_Persist.stLIC101Cfg
    stPidRetain  : PL.ST_DeviceRetain;                // GVL_Persist.stLIC101Retain
    fbAlarms     : FB_StationAlarms;                  // GVL_Station.fbAlarms
    rOutBefore   : REAL;                              // выход LIC101 до события
    rMinSp       : REAL;                              // наименьшее общее задание частоты после события
    uiStep       : UINT;                              // шаг после события
END_VAR

(* ---- PidHandoverKeepsOutput.method.impl.st ---- *)
coUnit.TEST('StationCore_PidHandoverKeepsOutput_A7_A8');

StartPidTwoPumps(fbDut := fbDut, fbTime := fbTime, stCmd := stCmd, stCfgPersist := stCfgPersist,
                 stCfgLkg := stCfgLkg, stRetain := stRetain, fbPid := fbPid, stPidCmd := stPidCmd,
                 stPidCfg := stPidCfg, stPidRetain := stPidRetain, fbAlarms := fbAlarms, afbPump := afbPump,
                 itfEvents := fbSink);
AssertTrue(Condition := fbDut.stSts.eControlAct = E_ControlAct.LevelPid, Message := 'LevelPid before the event');
AssertTrue(Condition := fbDut.stSts.uiLeadPump = 1 AND afbPump[1].xRunning AND afbPump[2].xRunning
                        AND NOT afbPump[3].xRunning, Message := 'lead 1 and assist 2 running, 3 standby');
AssertTrue(Condition := (fbPid.stSts.stCommon.wStatus AND PL.GVL_Const.PID_STS_TRACKING) = 0,
           Message := 'PID controls before the event');
AssertTrue(Condition := fbPid.rOut_pct > 80.0 AND fbPid.rOut_pct < 98.0, Message := 'PID output high, below 98 %');
rOutBefore := fbPid.rOut_pct;

// ведущий 1 работает без остановки дольше tMaxContRun (4 ч)
afbPump[1].udiCurrentRunSeconds := TIME_TO_UDINT(stCfgLkg.tMaxContRun) / GVL_Const.STN_MS_PER_S + 1;
rMinSp := fbDut.rSpeedSp_pct;
FOR uiStep := 1 TO 120 DO
    Cycle(fbDut := fbDut, fbTime := fbTime, stCmd := stCmd, stCfgPersist := stCfgPersist, stCfgLkg := stCfgLkg,
          stRetain := stRetain, fbPid := fbPid, stPidCmd := stPidCmd, stPidCfg := stPidCfg,
          stPidRetain := stPidRetain, fbAlarms := fbAlarms, afbPump := afbPump, tStep := T#100MS, uiSteps := 1,
          xPlant := TRUE);
    rMinSp := MIN(rMinSp, fbDut.rSpeedSp_pct);
END_FOR

AssertEquals_REAL(Expected := 3.0, Actual := fbSink.ValueOf(eFind := E_StationEvent.ContRunHandover), Delta := 0.0,
                  Message := 'event 101007 with pump 3');
AssertTrue(Condition := fbDut.axRun[2] AND fbDut.axRun[3] AND NOT fbDut.axRun[1],
           Message := 'pump 1 released after the overlap');
AssertEquals_UINT(Expected := 3, Actual := fbDut.stSts.uiLeadPump, Message := 'replacement 3 becomes lead');
AssertTrue(Condition := fbDut.stSts.eControlAct = E_ControlAct.LevelPid, Message := 'still LevelPid');
AssertTrue(Condition := (fbPid.stSts.stCommon.wStatus AND PL.GVL_Const.PID_STS_TRACKING) = 0,
           Message := 'PID controls via the new lead');
AssertTrue(Condition := rMinSp >= rOutBefore - 2.0, Message := 'speed setpoint did not collapse');
AssertEquals_REAL(Expected := rOutBefore, Actual := fbPid.rOut_pct, Delta := 5.0,
                  Message := 'PID output near the previous one');
AssertEquals_REAL(Expected := rOutBefore, Actual := afbPump[2].rSpeedRef, Delta := 5.0,
                  Message := 'pump 2 speed near the previous output');
AssertEquals_REAL(Expected := rOutBefore, Actual := afbPump[3].rSpeedRef, Delta := 5.0,
                  Message := 'pump 3 speed near the previous output');
AssertEquals_UINT(Expected := 2, Actual := fbDut.stSts.uiPumpsRunning, Message := 'two pumps running');

coUnit.TEST_FINISHED();

(* ---- PidLeadFaultKeepsOutput.method.decl.st ---- *)
// 04 §7.3, §9, PMI-13 в режиме ПИД: авария ПЧ ведущего при двух работающих насосах — подпорный 2 становится
// ведущим, резервный 3 пускается в том же цикле, а выход LIC101 и частота насосов не проваливаются: в цикле отказа
// ПИД держит свой выход, а не следует за заданием 0 отказавшего ПЧ (дефект, найденный на рантайме при записи тренда)
METHOD PRIVATE PidLeadFaultKeepsOutput
VAR
    fbDut        : FB_StationCore;                    // ФБ под тестом
    fbTime       : PL.FB_FakeTime;                    // подменное время, старт 1 ч
    fbSink       : FB_FakeEventSink;                  // подменный журнал
    afbPump      : ARRAY[1..3] OF FB_FakeMotorVfd;    // подменные насосы: доступны, Auto, стоят
    stCmd        : ST_StationCmd;                     // GVL_Station.stStationCmd
    stCfgPersist : ST_StationCfg;                     // GVL_Persist.stStationCfg
    stCfgLkg     : ST_StationCfg;                     // GVL_Station.stCfgLkg
    stRetain     : ST_StationRetain;                  // GVL_Persist.stStationRetain
    fbPid        : PL.FB_PID;                         // GVL_Station.fbLIC101
    stPidCmd     : PL.ST_PidCmd;                      // GVL_Station.stLIC101Cmd
    stPidCfg     : PL.ST_PidCfg;                      // GVL_Persist.stLIC101Cfg
    stPidRetain  : PL.ST_DeviceRetain;                // GVL_Persist.stLIC101Retain
    fbAlarms     : FB_StationAlarms;                  // GVL_Station.fbAlarms
    rOutBefore   : REAL;                              // выход LIC101 до события
    rMinSp       : REAL;                              // наименьшее общее задание частоты после события
    uiStep       : UINT;                              // шаг после события
END_VAR

(* ---- PidLeadFaultKeepsOutput.method.impl.st ---- *)
coUnit.TEST('StationCore_PidLeadFaultKeepsOutput_A7_A9_PMI13');

StartPidTwoPumps(fbDut := fbDut, fbTime := fbTime, stCmd := stCmd, stCfgPersist := stCfgPersist,
                 stCfgLkg := stCfgLkg, stRetain := stRetain, fbPid := fbPid, stPidCmd := stPidCmd,
                 stPidCfg := stPidCfg, stPidRetain := stPidRetain, fbAlarms := fbAlarms, afbPump := afbPump,
                 itfEvents := fbSink);
AssertTrue(Condition := fbDut.stSts.eControlAct = E_ControlAct.LevelPid, Message := 'LevelPid before the event');
AssertTrue(Condition := fbDut.stSts.uiLeadPump = 1 AND afbPump[1].xRunning AND afbPump[2].xRunning
                        AND NOT afbPump[3].xRunning, Message := 'lead 1 and assist 2 running, 3 standby');
AssertTrue(Condition := (fbPid.stSts.stCommon.wStatus AND PL.GVL_Const.PID_STS_TRACKING) = 0,
           Message := 'PID controls before the event');
AssertTrue(Condition := fbPid.rOut_pct > 80.0 AND fbPid.rOut_pct < 98.0, Message := 'PID output high, below 98 %');
rOutBefore := fbPid.rOut_pct;

// авария ПЧ ведущего (USAGE §3): устройство останавливает насос, задание на ПЧ 0, насос недоступен
afbPump[1].xFault := TRUE;
afbPump[1].xRunning := FALSE;
afbPump[1].xSpeedAuto := FALSE;
afbPump[1].rSpeedRef := 0.0;
afbPump[1].rSpeedAct := 0.0;
Cycle(fbDut := fbDut, fbTime := fbTime, stCmd := stCmd, stCfgPersist := stCfgPersist, stCfgLkg := stCfgLkg,
      stRetain := stRetain, fbPid := fbPid, stPidCmd := stPidCmd, stPidCfg := stPidCfg,
      stPidRetain := stPidRetain, fbAlarms := fbAlarms, afbPump := afbPump, tStep := T#100MS, uiSteps := 1,
      xPlant := TRUE);

AssertTrue(Condition := fbDut.axRun[2] AND fbDut.axRun[3] AND NOT fbDut.axRun[1],
           Message := 'faulted lead released, standby 3 requested in the same cycle');
AssertEquals_UINT(Expected := 2, Actual := fbDut.stSts.uiLeadPump, Message := 'assist 2 becomes lead');
AssertEquals_REAL(Expected := rOutBefore, Actual := fbDut.rSpeedSp_pct, Delta := 0.5,
                  Message := 'fault cycle: speed setpoint keeps the PID output');
rMinSp := fbDut.rSpeedSp_pct;
FOR uiStep := 1 TO 30 DO
    Cycle(fbDut := fbDut, fbTime := fbTime, stCmd := stCmd, stCfgPersist := stCfgPersist, stCfgLkg := stCfgLkg,
          stRetain := stRetain, fbPid := fbPid, stPidCmd := stPidCmd, stPidCfg := stPidCfg,
          stPidRetain := stPidRetain, fbAlarms := fbAlarms, afbPump := afbPump, tStep := T#100MS, uiSteps := 1,
          xPlant := TRUE);
    rMinSp := MIN(rMinSp, fbDut.rSpeedSp_pct);
END_FOR

AssertTrue(Condition := fbDut.stSts.eControlAct = E_ControlAct.LevelPid, Message := 'still LevelPid');
AssertTrue(Condition := (fbPid.stSts.stCommon.wStatus AND PL.GVL_Const.PID_STS_TRACKING) = 0,
           Message := 'PID controls via the new lead');
AssertTrue(Condition := rMinSp >= rOutBefore - 2.0, Message := 'speed setpoint did not collapse');
AssertEquals_REAL(Expected := rOutBefore, Actual := fbPid.rOut_pct, Delta := 5.0,
                  Message := 'PID output near the previous one');
AssertEquals_REAL(Expected := rOutBefore, Actual := afbPump[2].rSpeedRef, Delta := 5.0,
                  Message := 'pump 2 speed near the previous output');
AssertEquals_REAL(Expected := rOutBefore, Actual := afbPump[3].rSpeedRef, Delta := 5.0,
                  Message := 'pump 3 speed near the previous output');
AssertEquals_UINT(Expected := 2, Actual := fbDut.stSts.uiPumpsRunning, Message := 'two pumps running');

coUnit.TEST_FINISHED();

(* ---- PidLeadTripKeepsOutput.method.decl.st ---- *)
// 04 §7.3, §9.1, §10.4, PMI-16 в режиме ПИД: перегрев обмотки ведущего (блокировка станции) при двух работающих
// насосах — устройство останавливает насос в цикле блокировки, роль передаётся в следующем; выход LIC101 и частота
// насосов не проваливаются: ПИД не следует за заданием 0 остановленного блокировкой ПЧ. Недогрузка (10.3) приходит
// через ту же блокировку станции wInterlock
METHOD PRIVATE PidLeadTripKeepsOutput
VAR
    fbDut        : FB_StationCore;                    // ФБ под тестом
    fbTime       : PL.FB_FakeTime;                    // подменное время, старт 1 ч
    fbSink       : FB_FakeEventSink;                  // подменный журнал
    afbPump      : ARRAY[1..3] OF FB_FakeMotorVfd;    // подменные насосы: доступны, Auto, стоят
    stCmd        : ST_StationCmd;                     // GVL_Station.stStationCmd
    stCfgPersist : ST_StationCfg;                     // GVL_Persist.stStationCfg
    stCfgLkg     : ST_StationCfg;                     // GVL_Station.stCfgLkg
    stRetain     : ST_StationRetain;                  // GVL_Persist.stStationRetain
    fbPid        : PL.FB_PID;                         // GVL_Station.fbLIC101
    stPidCmd     : PL.ST_PidCmd;                      // GVL_Station.stLIC101Cmd
    stPidCfg     : PL.ST_PidCfg;                      // GVL_Persist.stLIC101Cfg
    stPidRetain  : PL.ST_DeviceRetain;                // GVL_Persist.stLIC101Retain
    fbAlarms     : FB_StationAlarms;                  // GVL_Station.fbAlarms
    rOutBefore   : REAL;                              // выход LIC101 до события
    rMinSp       : REAL;                              // наименьшее общее задание частоты после события
    uiStep       : UINT;                              // шаг после события
END_VAR

(* ---- PidLeadTripKeepsOutput.method.impl.st ---- *)
coUnit.TEST('StationCore_PidLeadTripKeepsOutput_A7_A9_A10_PMI16');

StartPidTwoPumps(fbDut := fbDut, fbTime := fbTime, stCmd := stCmd, stCfgPersist := stCfgPersist,
                 stCfgLkg := stCfgLkg, stRetain := stRetain, fbPid := fbPid, stPidCmd := stPidCmd,
                 stPidCfg := stPidCfg, stPidRetain := stPidRetain, fbAlarms := fbAlarms, afbPump := afbPump,
                 itfEvents := fbSink);
AssertTrue(Condition := fbDut.stSts.eControlAct = E_ControlAct.LevelPid, Message := 'LevelPid before the event');
AssertTrue(Condition := fbDut.stSts.uiLeadPump = 1 AND afbPump[1].xRunning AND afbPump[2].xRunning
                        AND NOT afbPump[3].xRunning, Message := 'lead 1 and assist 2 running, 3 standby');
AssertTrue(Condition := (fbPid.stSts.stCommon.wStatus AND PL.GVL_Const.PID_STS_TRACKING) = 0,
           Message := 'PID controls before the event');
AssertTrue(Condition := fbPid.rOut_pct > 80.0 AND fbPid.rOut_pct < 98.0, Message := 'PID output high, below 98 %');
rOutBefore := fbPid.rOut_pct;

// TS112: блокировка станции в этом цикле
fbDut.axOverheat[1] := TRUE;
Cycle(fbDut := fbDut, fbTime := fbTime, stCmd := stCmd, stCfgPersist := stCfgPersist, stCfgLkg := stCfgLkg,
      stRetain := stRetain, fbPid := fbPid, stPidCmd := stPidCmd, stPidCfg := stPidCfg,
      stPidRetain := stPidRetain, fbAlarms := fbAlarms, afbPump := afbPump, tStep := T#100MS, uiSteps := 1,
      xPlant := TRUE);

AssertTrue(Condition := (fbDut.awInterlock[1] AND GVL_Const.KNS_ILK_OVERHEAT) <> 0, Message := 'overheat interlock');
// устройство выполнило блокировку: насос недоступен и останавливается, задание на ПЧ 0; авария ПЧ — позже
afbPump[1].xAvailable := FALSE;
afbPump[1].xRunning := FALSE;
afbPump[1].xSpeedAuto := FALSE;
afbPump[1].rSpeedRef := 0.0;
afbPump[1].rSpeedAct := 0.0;
rMinSp := fbDut.rSpeedSp_pct;
FOR uiStep := 1 TO 30 DO
    Cycle(fbDut := fbDut, fbTime := fbTime, stCmd := stCmd, stCfgPersist := stCfgPersist, stCfgLkg := stCfgLkg,
          stRetain := stRetain, fbPid := fbPid, stPidCmd := stPidCmd, stPidCfg := stPidCfg,
          stPidRetain := stPidRetain, fbAlarms := fbAlarms, afbPump := afbPump, tStep := T#100MS, uiSteps := 1,
          xPlant := TRUE);
    rMinSp := MIN(rMinSp, fbDut.rSpeedSp_pct);
END_FOR

AssertTrue(Condition := fbDut.axRun[2] AND fbDut.axRun[3] AND NOT fbDut.axRun[1],
           Message := 'tripped lead released, standby 3 requested');
AssertEquals_UINT(Expected := 2, Actual := fbDut.stSts.uiLeadPump, Message := 'assist 2 becomes lead');
AssertTrue(Condition := fbDut.stSts.eControlAct = E_ControlAct.LevelPid, Message := 'still LevelPid');
AssertTrue(Condition := (fbPid.stSts.stCommon.wStatus AND PL.GVL_Const.PID_STS_TRACKING) = 0,
           Message := 'PID controls via the new lead');
AssertTrue(Condition := rMinSp >= rOutBefore - 2.0, Message := 'speed setpoint did not collapse');
AssertEquals_REAL(Expected := rOutBefore, Actual := fbPid.rOut_pct, Delta := 5.0,
                  Message := 'PID output near the previous one');
AssertEquals_REAL(Expected := rOutBefore, Actual := afbPump[2].rSpeedRef, Delta := 5.0,
                  Message := 'pump 2 speed near the previous output');
AssertEquals_REAL(Expected := rOutBefore, Actual := afbPump[3].rSpeedRef, Delta := 5.0,
                  Message := 'pump 3 speed near the previous output');
AssertEquals_UINT(Expected := 2, Actual := fbDut.stSts.uiPumpsRunning, Message := 'two pumps running');

coUnit.TEST_FINISHED();

(* ---- PlcStartLogsEventAndDelaysRequests.method.decl.st ---- *)
// 04 §13.3, PMI-01, PMI-35: старт приложения — событие 101015 первым, последовательный пуск: до tPlcStart запросов
// нет даже при уровне выше пуска, затем ведущий
METHOD PRIVATE PlcStartLogsEventAndDelaysRequests
VAR
    fbDut        : FB_StationCore;                    // ФБ под тестом
    fbTime       : PL.FB_FakeTime;                    // подменное время, старт 1 ч
    fbSink       : FB_FakeEventSink;                  // подменный журнал
    afbPump      : ARRAY[1..3] OF FB_FakeMotorVfd;    // подменные насосы: доступны, Auto, стоят
    stCmd        : ST_StationCmd;                     // GVL_Station.stStationCmd
    stCfgPersist : ST_StationCfg;                     // GVL_Persist.stStationCfg
    stCfgLkg     : ST_StationCfg;                     // GVL_Station.stCfgLkg
    stRetain     : ST_StationRetain;                  // GVL_Persist.stStationRetain
    fbPid        : PL.FB_PID;                         // GVL_Station.fbLIC101
    stPidCmd     : PL.ST_PidCmd;                      // GVL_Station.stLIC101Cmd
    stPidCfg     : PL.ST_PidCfg;                      // GVL_Persist.stLIC101Cfg
    stPidRetain  : PL.ST_DeviceRetain;                // GVL_Persist.stLIC101Retain
    fbAlarms     : FB_StationAlarms;                  // GVL_Station.fbAlarms
END_VAR

(* ---- PowerLostSuppressesLackNoresAts.method.decl.st ---- *)
// 04 §13.1, PMI-33: нет напряжения — PowerLost, запросов нет; KNS1.NORES, KNS1.LACK, KNS1.ATS подавлены по условию
METHOD PRIVATE PowerLostSuppressesLackNoresAts
VAR
    fbDut        : FB_StationCore;                    // ФБ под тестом
    fbTime       : PL.FB_FakeTime;                    // подменное время, старт 1 ч
    fbSink       : FB_FakeEventSink;                  // подменный журнал
    afbPump      : ARRAY[1..3] OF FB_FakeMotorVfd;    // подменные насосы: доступны, Auto, стоят
    stCmd        : ST_StationCmd;                     // GVL_Station.stStationCmd
    stCfgPersist : ST_StationCfg;                     // GVL_Persist.stStationCfg
    stCfgLkg     : ST_StationCfg;                     // GVL_Station.stCfgLkg
    stRetain     : ST_StationRetain;                  // GVL_Persist.stStationRetain
    fbPid        : PL.FB_PID;                         // GVL_Station.fbLIC101
    stPidCmd     : PL.ST_PidCmd;                      // GVL_Station.stLIC101Cmd
    stPidCfg     : PL.ST_PidCfg;                      // GVL_Persist.stLIC101Cfg
    stPidRetain  : PL.ST_DeviceRetain;                // GVL_Persist.stLIC101Retain
    fbAlarms     : FB_StationAlarms;                  // GVL_Station.fbAlarms
    itfAlm       : PL.I_Alarm;                        // тревога через интерфейс
END_VAR

(* ---- ResetButtonEdgeResetsAndLogs.method.decl.st ---- *)
// 04 §14, PMI-36 шаг 7: фронт HS501 — общий сброс один раз (Reset() устройств, фиксации насосов), событие 101016
// со значением 1
METHOD PRIVATE ResetButtonEdgeResetsAndLogs
VAR
    fbDut        : FB_StationCore;                    // ФБ под тестом
    fbTime       : PL.FB_FakeTime;                    // подменное время, старт 1 ч
    fbSink       : FB_FakeEventSink;                  // подменный журнал
    afbPump      : ARRAY[1..3] OF FB_FakeMotorVfd;    // подменные насосы: доступны, Auto, стоят
    stCmd        : ST_StationCmd;                     // GVL_Station.stStationCmd
    stCfgPersist : ST_StationCfg;                     // GVL_Persist.stStationCfg
    stCfgLkg     : ST_StationCfg;                     // GVL_Station.stCfgLkg
    stRetain     : ST_StationRetain;                  // GVL_Persist.stStationRetain
    fbPid        : PL.FB_PID;                         // GVL_Station.fbLIC101
    stPidCmd     : PL.ST_PidCmd;                      // GVL_Station.stLIC101Cmd
    stPidCfg     : PL.ST_PidCfg;                      // GVL_Persist.stLIC101Cfg
    stPidRetain  : PL.ST_DeviceRetain;                // GVL_Persist.stLIC101Retain
    fbAlarms     : FB_StationAlarms;                  // GVL_Station.fbAlarms
END_VAR

(* ---- RestartSequencesEmergencyPumps.method.decl.st ---- *)
// 04 §13.2, §10.2, PMI-34: питание восстановлено при аварийно высоком уровне — последовательный пуск охватывает все
// насосы аварийного режима (ведущий, подпорный, остальные), каждый следующий — через tSeqStep после ОС предыдущего,
// на полной частоте. Третий насос не обходит tSeqStep интервалом tStagger
METHOD PRIVATE RestartSequencesEmergencyPumps
VAR
    fbDut        : FB_StationCore;                    // ФБ под тестом
    fbTime       : PL.FB_FakeTime;                    // подменное время, старт 1 ч
    fbSink       : FB_FakeEventSink;                  // подменный журнал
    afbPump      : ARRAY[1..3] OF FB_FakeMotorVfd;    // подменные насосы: доступны, Auto, стоят
    stCmd        : ST_StationCmd;                     // GVL_Station.stStationCmd
    stCfgPersist : ST_StationCfg;                     // GVL_Persist.stStationCfg
    stCfgLkg     : ST_StationCfg;                     // GVL_Station.stCfgLkg
    stRetain     : ST_StationRetain;                  // GVL_Persist.stStationRetain
    fbPid        : PL.FB_PID;                         // GVL_Station.fbLIC101
    stPidCmd     : PL.ST_PidCmd;                      // GVL_Station.stLIC101Cmd
    stPidCfg     : PL.ST_PidCfg;                      // GVL_Persist.stLIC101Cfg
    stPidRetain  : PL.ST_DeviceRetain;                // GVL_Persist.stLIC101Retain
    fbAlarms     : FB_StationAlarms;                  // GVL_Station.fbAlarms
    uiIdx        : UINT;                              // насос
    uiReq        : UINT;                              // выданных запросов
END_VAR

(* ---- RestartSequencesEmergencyPumps.method.impl.st ---- *)
coUnit.TEST('StationCore_RestartSequencesEmergencyPumps_A10_A13_PMI34');

stPidCfg := GVL_StationDefaults.stLIC101Cfg;
stRetain.eMode := E_StationMode.Auto;
stCfgPersist.rStepSpeed_pct := 80.0;                  // частота ступенчатого отличается от полной
fbDut.aitfPump[1] := afbPump[1];
fbDut.aitfPump[2] := afbPump[2];
fbDut.aitfPump[3] := afbPump[3];
fbDut.axCommOk[1] := TRUE;
fbDut.axCommOk[2] := TRUE;
fbDut.axCommOk[3] := TRUE;
fbDut.itfEvents := fbSink;
fbDut.rLevel_m := 1.2;
fbDut.xLevelValid := TRUE;
fbDut.eLevelNe107 := PL.E_Ne107Status.Good;
fbDut.rLvlL_m := 0.8;
fbDut.rLvlH_m := 3.5;
fbDut.xPowerOk := TRUE;
Cycle(fbDut := fbDut, fbTime := fbTime, stCmd := stCmd, stCfgPersist := stCfgPersist, stCfgLkg := stCfgLkg,
      stRetain := stRetain, fbPid := fbPid, stPidCmd := stPidCmd, stPidCfg := stPidCfg,
      stPidRetain := stPidRetain, fbAlarms := fbAlarms, afbPump := afbPump, tStep := T#100MS, uiSteps := 110,
      xPlant := TRUE);

// пропадание напряжения: насосы недоступны; за время без питания уровень дошёл до HH и LS102
fbDut.xPowerOk := FALSE;
FOR uiIdx := 1 TO 3 DO
    afbPump[uiIdx].xAvailable := FALSE;
END_FOR
fbDut.rLevel_m := 4.1;
fbDut.xLevelH := TRUE;
fbDut.xLevelHH := TRUE;
fbDut.xFloatHigh := TRUE;
Cycle(fbDut := fbDut, fbTime := fbTime, stCmd := stCmd, stCfgPersist := stCfgPersist, stCfgLkg := stCfgLkg,
      stRetain := stRetain, fbPid := fbPid, stPidCmd := stPidCmd, stPidCfg := stPidCfg,
      stPidRetain := stPidRetain, fbAlarms := fbAlarms, afbPump := afbPump, tStep := T#100MS, uiSteps := 50,
      xPlant := TRUE);

AssertTrue(Condition := fbDut.stSts.eControlAct = E_ControlAct.PowerLost, Message := 'PowerLost');
// восстановление: задержка tPwrRestart 10 с, затем шаги по tSeqStep 15 с
fbDut.xPowerOk := TRUE;
FOR uiIdx := 1 TO 3 DO
    afbPump[uiIdx].xAvailable := TRUE;
END_FOR
Cycle(fbDut := fbDut, fbTime := fbTime, stCmd := stCmd, stCfgPersist := stCfgPersist, stCfgLkg := stCfgLkg,
      stRetain := stRetain, fbPid := fbPid, stPidCmd := stPidCmd, stPidCfg := stPidCfg,
      stPidRetain := stPidRetain, fbAlarms := fbAlarms, afbPump := afbPump, tStep := T#100MS, uiSteps := 105,
      xPlant := TRUE);

uiReq := BOOL_TO_UINT(fbDut.axRun[1]) + BOOL_TO_UINT(fbDut.axRun[2]) + BOOL_TO_UINT(fbDut.axRun[3]);
AssertTrue(Condition := fbDut.stSts.eControlAct = E_ControlAct.Restart, Message := 'Restart: step 1');
AssertEquals_UINT(Expected := 1, Actual := uiReq, Message := 'step 1: one request');
AssertEquals_UINT(Expected := 3, Actual := fbDut.stSts.uiPumpsRequired, Message := 'emergency: all pumps required');
AssertEquals_REAL(Expected := 100.0, Actual := fbDut.rSpeedSp_pct, Delta := 0.0, Message := 'emergency: full speed');
Cycle(fbDut := fbDut, fbTime := fbTime, stCmd := stCmd, stCfgPersist := stCfgPersist, stCfgLkg := stCfgLkg,
      stRetain := stRetain, fbPid := fbPid, stPidCmd := stPidCmd, stPidCfg := stPidCfg,
      stPidRetain := stPidRetain, fbAlarms := fbAlarms, afbPump := afbPump, tStep := T#100MS, uiSteps := 245,
      xPlant := TRUE);

uiReq := BOOL_TO_UINT(fbDut.axRun[1]) + BOOL_TO_UINT(fbDut.axRun[2]) + BOOL_TO_UINT(fbDut.axRun[3]);
AssertTrue(Condition := fbDut.stSts.eControlAct = E_ControlAct.Restart, Message := 'Restart: step 2');
AssertEquals_UINT(Expected := 2, Actual := uiReq, Message := 'step 2: third pump waits for tSeqStep');
Cycle(fbDut := fbDut, fbTime := fbTime, stCmd := stCmd, stCfgPersist := stCfgPersist, stCfgLkg := stCfgLkg,
      stRetain := stRetain, fbPid := fbPid, stPidCmd := stPidCmd, stPidCfg := stPidCfg,
      stPidRetain := stPidRetain, fbAlarms := fbAlarms, afbPump := afbPump, tStep := T#100MS, uiSteps := 70,
      xPlant := TRUE);

AssertTrue(Condition := fbDut.axRun[1] AND fbDut.axRun[2] AND fbDut.axRun[3], Message := 'step 3: all requested');
AssertTrue(Condition := fbDut.stSts.eControlAct = E_ControlAct.Emergency, Message := 'sequence done: Emergency');
AssertEquals_REAL(Expected := 3.0, Actual := fbSink.ValueOf(eFind := E_StationEvent.RestartDone), Delta := 0.0,
                  Message := 'event 101010: three starts');

coUnit.TEST_FINISHED();

(* ---- RestoredInvalidLkgFallsBackToDefaults.method.decl.st ---- *)
// 04 §18.3: сохранённая копия LKG проверяется при старте как записанные уставки. Неверная копия (задание 2,6 м
// вне пределов LIC101 — например, после смены пределов задания) при неверных записанных уставках не
// применяется: станция работает по уставкам проекта, копия заменяется ими
METHOD PRIVATE RestoredInvalidLkgFallsBackToDefaults
VAR
    fbDut          : FB_StationCore;                  // ФБ под тестом (первый вызов — старт ПЛК)
    fbTime         : PL.FB_FakeTime;                  // подменное время, старт 1 ч
    fbSink         : FB_FakeEventSink;                // подменный журнал
    afbPump        : ARRAY[1..3] OF FB_FakeMotorVfd;  // подменные насосы: доступны, Auto, стоят
    stCmd          : ST_StationCmd;                   // GVL_Station.stStationCmd
    stCfgPersist   : ST_StationCfg;                   // GVL_Persist.stStationCfg
    stCfgLkg       : ST_StationCfg;                   // GVL_Station.stCfgLkg
    stCfgLkgRetain : ST_StationCfg;                   // GVL_Persist.stStationCfgLkg
    stRetain       : ST_StationRetain;                // GVL_Persist.stStationRetain
    fbPid          : PL.FB_PID;                       // GVL_Station.fbLIC101
    stPidCmd       : PL.ST_PidCmd;                    // GVL_Station.stLIC101Cmd
    stPidCfg       : PL.ST_PidCfg;                    // GVL_Persist.stLIC101Cfg
    stPidRetain    : PL.ST_DeviceRetain;              // GVL_Persist.stLIC101Retain
    fbAlarms       : FB_StationAlarms;                // GVL_Station.fbAlarms
    stDef          : ST_StationCfg;                   // уставки проекта (GVL_StationDefaults)
END_VAR

(* ---- RevertCfgRestoresLkg.method.decl.st ---- *)
// 04 §18.3, 08 §14 вопрос 2: xRevertCfg возвращает записанные уставки к действующей копии; событие 101017 со
// значением 0
METHOD PRIVATE RevertCfgRestoresLkg
VAR
    fbDut        : FB_StationCore;                    // ФБ под тестом
    fbTime       : PL.FB_FakeTime;                    // подменное время, старт 1 ч
    fbSink       : FB_FakeEventSink;                  // подменный журнал
    afbPump      : ARRAY[1..3] OF FB_FakeMotorVfd;    // подменные насосы: доступны, Auto, стоят
    stCmd        : ST_StationCmd;                     // GVL_Station.stStationCmd
    stCfgPersist : ST_StationCfg;                     // GVL_Persist.stStationCfg
    stCfgLkg     : ST_StationCfg;                     // GVL_Station.stCfgLkg
    stRetain     : ST_StationRetain;                  // GVL_Persist.stStationRetain
    fbPid        : PL.FB_PID;                         // GVL_Station.fbLIC101
    stPidCmd     : PL.ST_PidCmd;                      // GVL_Station.stLIC101Cmd
    stPidCfg     : PL.ST_PidCfg;                      // GVL_Persist.stLIC101Cfg
    stPidRetain  : PL.ST_DeviceRetain;                // GVL_Persist.stLIC101Retain
    fbAlarms     : FB_StationAlarms;                  // GVL_Station.fbAlarms
END_VAR

(* ---- SimulationAlarmAndFaultEvent.method.decl.st ---- *)
// ARCHITECTURE 4, PMI-01: имитация — KNS1.SIM, бит 11 wState, NE 107 C; рост счётчика инъекций — событие 101021
METHOD PRIVATE SimulationAlarmAndFaultEvent
VAR
    fbDut        : FB_StationCore;                    // ФБ под тестом
    fbTime       : PL.FB_FakeTime;                    // подменное время, старт 1 ч
    fbSink       : FB_FakeEventSink;                  // подменный журнал
    afbPump      : ARRAY[1..3] OF FB_FakeMotorVfd;    // подменные насосы: доступны, Auto, стоят
    stCmd        : ST_StationCmd;                     // GVL_Station.stStationCmd
    stCfgPersist : ST_StationCfg;                     // GVL_Persist.stStationCfg
    stCfgLkg     : ST_StationCfg;                     // GVL_Station.stCfgLkg
    stRetain     : ST_StationRetain;                  // GVL_Persist.stStationRetain
    fbPid        : PL.FB_PID;                         // GVL_Station.fbLIC101
    stPidCmd     : PL.ST_PidCmd;                      // GVL_Station.stLIC101Cmd
    stPidCfg     : PL.ST_PidCfg;                      // GVL_Persist.stLIC101Cfg
    stPidRetain  : PL.ST_DeviceRetain;                // GVL_Persist.stLIC101Retain
    fbAlarms     : FB_StationAlarms;                  // GVL_Station.fbAlarms
END_VAR

(* ---- StartPidTwoPumps.method.decl.st ---- *)
// Помощник: способ ПИД, LIC101 в Auto, старт ПЛК; пуск ведущего 1 по уровню 1,7 м, затем уровень 2,45 м —
// подпорный 2 по уровню (04 §7.2), выход ПИД около 90 % (подменные насосы следуют общему заданию частоты без
// минимальной частоты и рампы); после пуска подпорного выдерживается tStagger, чтобы резервный мог пуститься сразу
METHOD PRIVATE StartPidTwoPumps
VAR_IN_OUT
    fbDut        : FB_StationCore;                    // ФБ под тестом
    fbTime       : PL.FB_FakeTime;                    // подменное время
    stCmd        : ST_StationCmd;                     // команды
    stCfgPersist : ST_StationCfg;                     // записанные уставки
    stCfgLkg     : ST_StationCfg;                     // действующая копия
    stRetain     : ST_StationRetain;                  // режим, способ
    fbPid        : PL.FB_PID;                         // LIC101
    stPidCmd     : PL.ST_PidCmd;                      // команды LIC101
    stPidCfg     : PL.ST_PidCfg;                      // уставки LIC101
    stPidRetain  : PL.ST_DeviceRetain;                // режим LIC101
    fbAlarms     : FB_StationAlarms;                  // тревоги станции
    afbPump      : ARRAY[1..3] OF FB_FakeMotorVfd;    // подменные насосы
END_VAR
VAR_INPUT
    itfEvents : I_StationEventSink;                   // подменный журнал
END_VAR

(* ---- StationDefaultsMatchTypeDefaults.method.decl.st ---- *)
// DESIGN 4.2: GVL_StationDefaults.stStationCfg совпадает с умолчаниями ST_StationCfg по всем параметрам, тревогам
// и резерву (сравнение полей — без байтов выравнивания ST_AlarmCfg); границы резерва — по константам
// STN_CFG_RESERVE_*
METHOD PRIVATE StationDefaultsMatchTypeDefaults
VAR
    fbDut   : FB_StationCore;           // метод сравнения уставок
    stDef   : ST_StationCfg;            // копия константы GVL_StationDefaults
    stType  : ST_StationCfg;            // умолчания типа
END_VAR

(* ---- StationStsSizeIs72.method.decl.st ---- *)
// 04 §19.3, DESIGN 3.1: ST_StationSts — только 16- и 32-битные поля, 72 байта (раскладка для OPC UA и MQTT)
METHOD PRIVATE StationStsSizeIs72
VAR
    stSts : ST_StationSts;              // проверяемая структура
END_VAR

(* ---- StepAlarmNoFlickerAfterPowerRestorePid.method.decl.st ---- *)
// 04 §7.4, §12, §13, §15, PMI-33, PMI-34: выбран ПИД, пропадание напряжения 30 с, восстановление. Пока нет
// напряжения, насосы недоступны и без связи (ПЧ без питания); после восстановления ПЧ ещё 2 с загружаются (связи
// нет). Последовательный пуск — штатный переходный режим: KNS1.STEP подавлена, загрузка ПЧ — не потеря связи
// (VFD-12), выдержка STN_PID_RECOVER не перезапускается. После последовательного пуска — сразу ПИД, STEP нет
METHOD PRIVATE StepAlarmNoFlickerAfterPowerRestorePid
VAR
    fbDut        : FB_StationCore;                    // ФБ под тестом
    fbTime       : PL.FB_FakeTime;                    // подменное время, старт 1 ч
    fbSink       : FB_FakeEventSink;                  // подменный журнал
    afbPump      : ARRAY[1..3] OF FB_FakeMotorVfd;    // подменные насосы: доступны, Auto, стоят
    stCmd        : ST_StationCmd;                     // GVL_Station.stStationCmd
    stCfgPersist : ST_StationCfg;                     // GVL_Persist.stStationCfg
    stCfgLkg     : ST_StationCfg;                     // GVL_Station.stCfgLkg
    stRetain     : ST_StationRetain;                  // GVL_Persist.stStationRetain
    fbPid        : PL.FB_PID;                         // GVL_Station.fbLIC101
    stPidCmd     : PL.ST_PidCmd;                      // GVL_Station.stLIC101Cmd
    stPidCfg     : PL.ST_PidCfg;                      // GVL_Persist.stLIC101Cfg
    stPidRetain  : PL.ST_DeviceRetain;                // GVL_Persist.stLIC101Retain
    fbAlarms     : FB_StationAlarms;                  // GVL_Station.fbAlarms
    itfStep      : PL.I_Alarm;                        // KNS1.STEP через интерфейс
    uiIdx        : UINT;                              // насос
    uiStep       : UINT;                              // шаг
    xFlicker     : BOOL;                              // STEP была неквитированной хотя бы в одном цикле
END_VAR

(* ---- StepAlarmNoFlickerAfterPowerRestorePid.method.impl.st ---- *)
coUnit.TEST('StationCore_StepAlarmNoFlickerAfterPowerRestorePid_A7_A12_A13_A15_PMI33_PMI34');

stPidCfg := GVL_StationDefaults.stLIC101Cfg;
stRetain.eMode := E_StationMode.Auto;
stRetain.eMethod := E_ControlMethod.LevelPid;
stPidRetain.eRemoteMode := PL.E_DeviceMode.Auto;
fbDut.aitfPump[1] := afbPump[1];
fbDut.aitfPump[2] := afbPump[2];
fbDut.aitfPump[3] := afbPump[3];
fbDut.axCommOk[1] := TRUE;
fbDut.axCommOk[2] := TRUE;
fbDut.axCommOk[3] := TRUE;
fbDut.itfEvents := fbSink;
fbDut.rLevel_m := 1.2;
fbDut.xLevelValid := TRUE;
fbDut.eLevelNe107 := PL.E_Ne107Status.Good;
fbDut.rLvlL_m := 0.8;
fbDut.rLvlH_m := 3.5;
fbDut.xPowerOk := TRUE;
Cycle(fbDut := fbDut, fbTime := fbTime, stCmd := stCmd, stCfgPersist := stCfgPersist, stCfgLkg := stCfgLkg,
      stRetain := stRetain, fbPid := fbPid, stPidCmd := stPidCmd, stPidCfg := stPidCfg,
      stPidRetain := stPidRetain, fbAlarms := fbAlarms, afbPump := afbPump, tStep := T#100MS, uiSteps := 110,
      xPlant := TRUE);

AssertTrue(Condition := fbDut.stSts.eControlAct = E_ControlAct.LevelPid, Message := 'LevelPid before power loss');
// нет напряжения: со следующего цикла насосы недоступны и без связи (ПЧ без питания)
fbDut.xPowerOk := FALSE;
Cycle(fbDut := fbDut, fbTime := fbTime, stCmd := stCmd, stCfgPersist := stCfgPersist, stCfgLkg := stCfgLkg,
      stRetain := stRetain, fbPid := fbPid, stPidCmd := stPidCmd, stPidCfg := stPidCfg,
      stPidRetain := stPidRetain, fbAlarms := fbAlarms, afbPump := afbPump, tStep := T#100MS, uiSteps := 1,
      xPlant := TRUE);
FOR uiIdx := 1 TO 3 DO
    afbPump[uiIdx].xAvailable := FALSE;
    fbDut.axCommOk[uiIdx] := FALSE;
END_FOR
Cycle(fbDut := fbDut, fbTime := fbTime, stCmd := stCmd, stCfgPersist := stCfgPersist, stCfgLkg := stCfgLkg,
      stRetain := stRetain, fbPid := fbPid, stPidCmd := stPidCmd, stPidCfg := stPidCfg,
      stPidRetain := stPidRetain, fbAlarms := fbAlarms, afbPump := afbPump, tStep := T#100MS, uiSteps := 300,
      xPlant := TRUE);

AssertTrue(Condition := fbDut.stSts.eControlAct = E_ControlAct.PowerLost, Message := 'PowerLost');
itfStep := fbAlarms.GetAlarm(uiIndex := E_StationAlarm.STEP - 1);
AssertTrue(Condition := itfStep.State = PL.E_AlarmState.SuppressedByDesign, Message := 'PowerLost: STEP suppressed');
// напряжение восстановлено (ES301 подтвердил): насосы доступны циклом позже, ПЧ ещё 2 с загружаются
fbDut.xPowerOk := TRUE;
xFlicker := FALSE;
FOR uiStep := 1 TO 300 DO
    Cycle(fbDut := fbDut, fbTime := fbTime, stCmd := stCmd, stCfgPersist := stCfgPersist, stCfgLkg := stCfgLkg,
          stRetain := stRetain, fbPid := fbPid, stPidCmd := stPidCmd, stPidCfg := stPidCfg,
          stPidRetain := stPidRetain, fbAlarms := fbAlarms, afbPump := afbPump, tStep := T#100MS, uiSteps := 1,
          xPlant := TRUE);
    xFlicker := xFlicker OR (fbDut.stSts.wAlmUnack AND 16#0080) <> 0;
    IF uiStep = 1 THEN
        FOR uiIdx := 1 TO 3 DO
            afbPump[uiIdx].xAvailable := TRUE;
        END_FOR
    ELSIF uiStep = 21 THEN
        AssertTrue(Condition := fbDut.stSts.eControlAct = E_ControlAct.Restart, Message := 'sequential start');
        FOR uiIdx := 1 TO 3 DO
            fbDut.axCommOk[uiIdx] := TRUE;
        END_FOR
    END_IF
END_FOR

AssertFalse(Condition := xFlicker, Message := 'no unacked KNS1.STEP after power restore');
AssertTrue(Condition := itfStep.State = PL.E_AlarmState.Normal, Message := 'STEP normal');
AssertTrue(Condition := fbDut.stSts.eControlAct = E_ControlAct.LevelPid, Message := 'LevelPid 30 s after restore');
AssertEquals_WORD(Expected := 0, Actual := fbDut.stSts.wState AND GVL_Const.STN_ST_STEP_FALLBACK,
                  Message := 'wState: no step fallback bit');

coUnit.TEST_FINISHED();

(* ---- StepAlarmNoFlickerOnStartAndAutoEntry.method.decl.st ---- *)
// 04 §3.2, §7.4, §15, PMI-01, PMI-30: выбран ПИД — при старте ПЛК (LIC101 и насосы ещё не вызывались) и при
// переходе «Ручной» → «Автомат» (насосы ещё в Manual, доступных нет) готовность ПИД пару циклов ложна. Это не
// отказ: KNS1.STEP (Low) не появляется и не остаётся неквитированной (задержка появления тревоги)
METHOD PRIVATE StepAlarmNoFlickerOnStartAndAutoEntry
VAR
    fbDut        : FB_StationCore;                    // ФБ под тестом
    fbTime       : PL.FB_FakeTime;                    // подменное время, старт 1 ч
    fbSink       : FB_FakeEventSink;                  // подменный журнал
    afbPump      : ARRAY[1..3] OF FB_FakeMotorVfd;    // подменные насосы: доступны, Auto, стоят
    stCmd        : ST_StationCmd;                     // GVL_Station.stStationCmd
    stCfgPersist : ST_StationCfg;                     // GVL_Persist.stStationCfg
    stCfgLkg     : ST_StationCfg;                     // GVL_Station.stCfgLkg
    stRetain     : ST_StationRetain;                  // GVL_Persist.stStationRetain
    fbPid        : PL.FB_PID;                         // GVL_Station.fbLIC101
    stPidCmd     : PL.ST_PidCmd;                      // GVL_Station.stLIC101Cmd
    stPidCfg     : PL.ST_PidCfg;                      // GVL_Persist.stLIC101Cfg
    stPidRetain  : PL.ST_DeviceRetain;                // GVL_Persist.stLIC101Retain
    fbAlarms     : FB_StationAlarms;                  // GVL_Station.fbAlarms
    uiIdx        : UINT;                              // насос
END_VAR

(* ---- StepAlarmNoFlickerOnStartAndAutoEntry.method.impl.st ---- *)
coUnit.TEST('StationCore_StepAlarmNoFlickerOnStartAndAutoEntry_A3_A7_A15_PMI01_PMI30');

stPidCfg := GVL_StationDefaults.stLIC101Cfg;
stRetain.eMode := E_StationMode.Auto;
fbDut.aitfPump[1] := afbPump[1];
fbDut.aitfPump[2] := afbPump[2];
fbDut.aitfPump[3] := afbPump[3];
fbDut.axCommOk[1] := TRUE;
fbDut.axCommOk[2] := TRUE;
fbDut.axCommOk[3] := TRUE;
fbDut.itfEvents := fbSink;
fbDut.rLevel_m := 1.2;
fbDut.xLevelValid := TRUE;
fbDut.eLevelNe107 := PL.E_Ne107Status.Good;
fbDut.rLvlL_m := 0.8;
fbDut.rLvlH_m := 3.5;
fbDut.xPowerOk := TRUE;

stRetain.eMethod := E_ControlMethod.LevelPid;
stPidRetain.eRemoteMode := PL.E_DeviceMode.Auto;
FOR uiIdx := 1 TO 3 DO
    afbPump[uiIdx].xFollowRequests := TRUE;
END_FOR
// старт ПЛК в «Автомате» с выбранным ПИД
Cycle(fbDut := fbDut, fbTime := fbTime, stCmd := stCmd, stCfgPersist := stCfgPersist, stCfgLkg := stCfgLkg,
      stRetain := stRetain, fbPid := fbPid, stPidCmd := stPidCmd, stPidCfg := stPidCfg,
      stPidRetain := stPidRetain, fbAlarms := fbAlarms, afbPump := afbPump, tStep := T#20MS, uiSteps := 600,
      xPlant := TRUE);

AssertTrue(Condition := fbDut.stSts.eControlAct = E_ControlAct.LevelPid, Message := 'start: LevelPid');
AssertEquals_WORD(Expected := 0, Actual := fbDut.stSts.wAlmUnack AND 16#0080, Message := 'start: no KNS1.STEP');
// «Ручной», насос Н1 пущен оператором
stCmd.xSetManual := TRUE;
Cycle(fbDut := fbDut, fbTime := fbTime, stCmd := stCmd, stCfgPersist := stCfgPersist, stCfgLkg := stCfgLkg,
      stRetain := stRetain, fbPid := fbPid, stPidCmd := stPidCmd, stPidCfg := stPidCfg,
      stPidRetain := stPidRetain, fbAlarms := fbAlarms, afbPump := afbPump, tStep := T#20MS, uiSteps := 5,
      xPlant := TRUE);

AssertTrue(Condition := afbPump[1].eMode = PL.E_DeviceMode.Manual, Message := 'pumps in Manual');
afbPump[1].xRunning := TRUE;
afbPump[1].rSpeedRef := 80.0;
afbPump[1].rSpeedAct := 80.0;
fbDut.rLevel_m := 1.5;
Cycle(fbDut := fbDut, fbTime := fbTime, stCmd := stCmd, stCfgPersist := stCfgPersist, stCfgLkg := stCfgLkg,
      stRetain := stRetain, fbPid := fbPid, stPidCmd := stPidCmd, stPidCfg := stPidCfg,
      stPidRetain := stPidRetain, fbAlarms := fbAlarms, afbPump := afbPump, tStep := T#20MS, uiSteps := 50,
      xPlant := TRUE);

// «Автомат»: насосы переходят в Auto в своём вызове
stCmd.xSetAuto := TRUE;
Cycle(fbDut := fbDut, fbTime := fbTime, stCmd := stCmd, stCfgPersist := stCfgPersist, stCfgLkg := stCfgLkg,
      stRetain := stRetain, fbPid := fbPid, stPidCmd := stPidCmd, stPidCfg := stPidCfg,
      stPidRetain := stPidRetain, fbAlarms := fbAlarms, afbPump := afbPump, tStep := T#20MS, uiSteps := 100,
      xPlant := TRUE);

AssertTrue(Condition := fbDut.stSts.eControlAct = E_ControlAct.LevelPid, Message := 'Auto entry: LevelPid');
AssertTrue(Condition := fbDut.axRun[1] AND afbPump[1].xRunning, Message := 'running pump adopted');
AssertEquals_WORD(Expected := 0, Actual := fbDut.stSts.wAlmUnack AND 16#0080, Message := 'Auto entry: no KNS1.STEP');

coUnit.TEST_FINISHED();

(* ---- StepFallbackSuppressedInEmergency.method.decl.st ---- *)
// 04 §7.4, §15: выбран ПИД, ПИД не готов (LIC101 в Manual) — ступенчатое и KNS1.STEP (после последовательного
// пуска старта ПЛК и своей выдержки 10 с); в аварийном режиме STEP подавлена
METHOD PRIVATE StepFallbackSuppressedInEmergency
VAR
    fbDut        : FB_StationCore;                    // ФБ под тестом
    fbTime       : PL.FB_FakeTime;                    // подменное время, старт 1 ч
    fbSink       : FB_FakeEventSink;                  // подменный журнал
    afbPump      : ARRAY[1..3] OF FB_FakeMotorVfd;    // подменные насосы: доступны, Auto, стоят
    stCmd        : ST_StationCmd;                     // GVL_Station.stStationCmd
    stCfgPersist : ST_StationCfg;                     // GVL_Persist.stStationCfg
    stCfgLkg     : ST_StationCfg;                     // GVL_Station.stCfgLkg
    stRetain     : ST_StationRetain;                  // GVL_Persist.stStationRetain
    fbPid        : PL.FB_PID;                         // GVL_Station.fbLIC101
    stPidCmd     : PL.ST_PidCmd;                      // GVL_Station.stLIC101Cmd
    stPidCfg     : PL.ST_PidCfg;                      // GVL_Persist.stLIC101Cfg
    stPidRetain  : PL.ST_DeviceRetain;                // GVL_Persist.stLIC101Retain
    fbAlarms     : FB_StationAlarms;                  // GVL_Station.fbAlarms
    itfAlm       : PL.I_Alarm;                        // тревога через интерфейс
END_VAR

(* ---- UnderloadTripInterlocksAndAts.method.decl.st ---- *)
// 04 §10.3, PMI-15: недогрузка ведущего — фиксация, KNS_ILK_UNDERLOAD, KNS1.UL1, АВР; сброс насоса снимает
// фиксацию
METHOD PRIVATE UnderloadTripInterlocksAndAts
VAR
    fbDut        : FB_StationCore;                    // ФБ под тестом
    fbTime       : PL.FB_FakeTime;                    // подменное время, старт 1 ч
    fbSink       : FB_FakeEventSink;                  // подменный журнал
    afbPump      : ARRAY[1..3] OF FB_FakeMotorVfd;    // подменные насосы: доступны, Auto, стоят
    stCmd        : ST_StationCmd;                     // GVL_Station.stStationCmd
    stCfgPersist : ST_StationCfg;                     // GVL_Persist.stStationCfg
    stCfgLkg     : ST_StationCfg;                     // GVL_Station.stCfgLkg
    stRetain     : ST_StationRetain;                  // GVL_Persist.stStationRetain
    fbPid        : PL.FB_PID;                         // GVL_Station.fbLIC101
    stPidCmd     : PL.ST_PidCmd;                      // GVL_Station.stLIC101Cmd
    stPidCfg     : PL.ST_PidCfg;                      // GVL_Persist.stLIC101Cfg
    stPidRetain  : PL.ST_DeviceRetain;                // GVL_Persist.stLIC101Retain
    fbAlarms     : FB_StationAlarms;                  // GVL_Station.fbAlarms
END_VAR

(* ---- VentilationAndAnnunciatorOutputs.method.decl.st ---- *)
// 04 §14, §17, PMI-36, PMI-38: выходы В1 и местной сигнализации — газ включает В1, пожар блокирует; новая High —
// сирена, активная High — K1 обесточено, бит 13 wState
METHOD PRIVATE VentilationAndAnnunciatorOutputs
VAR
    fbDut        : FB_StationCore;                    // ФБ под тестом
    fbTime       : PL.FB_FakeTime;                    // подменное время, старт 1 ч
    fbSink       : FB_FakeEventSink;                  // подменный журнал
    afbPump      : ARRAY[1..3] OF FB_FakeMotorVfd;    // подменные насосы: доступны, Auto, стоят
    stCmd        : ST_StationCmd;                     // GVL_Station.stStationCmd
    stCfgPersist : ST_StationCfg;                     // GVL_Persist.stStationCfg
    stCfgLkg     : ST_StationCfg;                     // GVL_Station.stCfgLkg
    stRetain     : ST_StationRetain;                  // GVL_Persist.stStationRetain
    fbPid        : PL.FB_PID;                         // GVL_Station.fbLIC101
    stPidCmd     : PL.ST_PidCmd;                      // GVL_Station.stLIC101Cmd
    stPidCfg     : PL.ST_PidCfg;                      // GVL_Persist.stLIC101Cfg
    stPidRetain  : PL.ST_DeviceRetain;                // GVL_Persist.stLIC101Retain
    fbAlarms     : FB_StationAlarms;                  // GVL_Station.fbAlarms
END_VAR
